(* IEC 61131-3 sources: daoli-st-library/DL_Motion (part 4) *)

(* ---- FC_DL_StackerMastSwayCalc.st ---- *)
(*
  DL Factory R83 | FC_DL_StackerMastSwayCalc
  功能：按加减速度与立柱高度估算堆垛机立柱顶部准静态摆幅与残余振荡稳定时间。
  开源溯源：无（clean-room 自研，依据公开工艺公式，来源=行业通用公式，许可证=MIT，借鉴点=公式结构）
  规则：R1-R21 全遵守
*)
FUNCTION FC_DL_StackerMastSwayCalc : REAL
VAR_INPUT
    fAccMs2    : REAL; // 行走加（减）速度 [m/s²] / Travel acceleration [m/s^2]
    fMastHM    : REAL; // 立柱有效悬臂高度 [m] / Effective mast cantilever height [m]
    fNatHz     : REAL; // 立柱一阶固有频率 [Hz] / First natural frequency of mast [Hz]
    fDampRatio : REAL; // 阻尼比（0.01~0.20）[-]/ Damping ratio [0.01..0.20]
    fDynFactor : REAL; // 悬臂动载放大系数（1.0~2.0）[-]/ Cantilever dynamic amplification [1.0..2.0]
END_VAR
VAR_OUTPUT
    fSwayMm  : REAL; // 立柱顶部准静态摆幅（单侧）[mm] / Quasi-static sway amplitude [mm]
    fSettleS : REAL; // 残余振荡衰减到 5% 的稳定时间 [s] / Settling time to 5 percent [s]
    fSwayDeg : REAL; // 立柱倾角（摆幅÷高度）[°] / Mast tilt angle [deg]
    xValid   : BOOL; // 计算有效性标志 / Calculation validity flag
END_VAR
VAR
    fAccG  : REAL; // 加速度折算重力倍数 [-] / Acceleration in g units
    fOmega : REAL; // 一阶圆频率 [rad/s] / First angular frequency [rad/s]
    cG     : REAL := 9.80665; // 标准重力加速度常量 [m/s²]，已引用（R19）/ Standard gravity [m/s^2]
END_VAR
// 出口预置：四出口统一预置（R256）
fSwayMm := 0.0; fSettleS := 0.0; fSwayDeg := 0.0; xValid := FALSE;
// 非有限拦截 + 量纲自检 + 分母零闸（R4/R20/R21）
IF NOT (fAccMs2 > -1.0E30 AND fAccMs2 < 1.0E30) OR NOT (fMastHM > -1.0E30 AND fMastHM < 1.0E30) OR NOT (fNatHz > -1.0E30 AND fNatHz < 1.0E30) OR NOT (fDampRatio > -1.0E30 AND fDampRatio < 1.0E30) OR NOT (fDynFactor > -1.0E30 AND fDynFactor < 1.0E30) OR fAccMs2 < 0.0 OR fMastHM <= 0.0 OR fNatHz <= 0.0 OR fDampRatio <= 0.0 OR fDynFactor <= 0.0 THEN
    FC_DL_StackerMastSwayCalc := -1.0; RETURN;  // 哨兵 -1：非有限或量纲越界 / Sentinel -1
END_IF
// 加速度折算：m/s² ÷ m/s² = 无量纲重力倍数（量纲自洽）
fAccG := fAccMs2 / cG;              // 重力倍数 [-] / Acceleration in g units
// 准静态摆幅：a/g × H × 动载放大，m × 1000 = mm（悬臂顶挠度正比于 aH/g）
fSwayMm := fAccG * fMastHM * fDynFactor * 1000.0;   // 单侧摆幅 [mm] / One-side sway [mm]
// 一阶圆频率：ω = 2πf，f 单位 Hz 得 rad/s（2π 为无量纲弧度量）
fOmega := 2.0 * 3.14159265358979 * fNatHz;          // 圆频率 [rad/s] / Angular frequency [rad/s]
// 稳定时间：4 ÷ (ζω) 近似衰减到 5%，分母显式零闸（R4/R21）
IF ABS(fDampRatio * fOmega) > 1.0E-9 THEN          // 阻尼×频率分母显式零闸 / Zero gate on damped frequency
    fSettleS := 4.0 / (fDampRatio * fOmega);        // 稳定时间 [s] / Settling time [s]
ELSE
    fSettleS := 0.0;                // 无阻尼不可估稳定时间，缺省零 / Undamped, default zero
END_IF
// 倾角：摆幅(mm) ÷ 高度(m×1000=mm) 得无量纲正切，×180/π 转度（小角近似）
fSwayDeg := (fSwayMm / (fMastHM * 1000.0)) * (180.0 / 3.14159265358979); // 倾角 [°] / Tilt [deg]
xValid := TRUE;                             // 链路有效 / Chain valid
FC_DL_StackerMastSwayCalc := fSwayMm;       // 返回单侧摆幅 [mm] / Return one-side sway [mm]
END_FUNCTION

(* ---- FC_DL_StanleySteerAngleCalc.st ---- *)
// FC_DL_StanleySteerAngleCalc v1.0.0
// 开源溯源：clean-room 自研（族 DL_Motion，ST 生态实测 0 命中，无外部代码引入）
(*
  功能: Stanley 前轮转角 δ = ψe + ATAN(k·e/(|v| + v_soft))，限幅 ±0.6 rad；
        软化速度负值归零，分母另设 1e-6 硬下限（双保险防除零）。
  邻件/码位: 与 FC_DL_AckermannSteerPairCalc 串联（转角→内外轮），与纯跟踪件互为替代律；
             16#0002_9205 = 域外或非有限拒收。
*)
FUNCTION FC_DL_StanleySteerAngleCalc : REAL
VAR_INPUT
    fHeadingErr : REAL := 0.0;      // 航向偏差 ψe [rad]，左正 / Heading error [rad]
    fCrossTrack : REAL := 0.0;      // 横向偏差 e [m]，左正 / Cross-track error [m]
    fSpeed      : REAL := 0.5;      // 车速 [m/s] / Vehicle speed [m/s]
    fGain       : REAL := 1.5;      // 横向增益 k [-]，域有限 / Cross-track gain [-]
    fSoft       : REAL := 0.2;      // 低速软化速度 [m/s]，负值取 0 / Softening speed [m/s]
END_VAR
VAR_OUTPUT
    fSteerAngle : REAL;             // 前轮转角 δ [rad]，限幅 ±0.6 / Steer angle [rad]
    bSaturated  : BOOL;             // 限幅命中标志 [-] / Saturation hit flag
    bValid      : BOOL;             // 结果有效回执 [-] / Result validity receipt
    uErrorId    : UDINT;            // 事件码，0 = 无事件 / Event code
END_VAR
VAR
    fSoftSafe : REAL := 0.0;        // 软化速度安全值 [m/s] / Sanitized softening speed [m/s]
    fDen      : REAL := 0.0;        // 分母 |v| + v_soft [m/s] / Denominator [m/s]
    fRaw      : REAL := 0.0;        // 未限幅转角 [rad] / Unsaturated angle [rad]
END_VAR
// 段 0：全路径出口安全缺省（转角零 = 直行）/ Safe defaults, zero angle means straight
fSteerAngle := 0.0;             // 转角缺省零 / Steer angle default zero
bSaturated := FALSE;            // 限幅标志预清 / Saturation preset clear
bValid := FALSE;                // 有效回执预清 / Validity preset clear
uErrorId := 16#0000;            // 事件码预清 / Event code preset clear
FC_DL_StanleySteerAngleCalc := 0.0;     // 返回值缺省零 / Return default zero
// 段 1：非有限闸（五入参全枚举）/ Non-finite gate over all inputs
IF (fHeadingErr <> fHeadingErr) OR (fCrossTrack <> fCrossTrack) OR (fSpeed <> fSpeed)
   OR (fGain <> fGain) OR (fSoft <> fSoft)
   OR (ABS(fHeadingErr) >= 3.0E38) OR (ABS(fCrossTrack) >= 3.0E38) OR (ABS(fSpeed) >= 3.0E38)
   OR (ABS(fGain) >= 3.0E38) OR (ABS(fSoft) >= 3.0E38) THEN
    uErrorId := 16#0002_9205;   // 入参非有限拒收 / Non-finite input reject
    RETURN;
END_IF
// 段 2：域闸（软化速度负值归零 + 分母硬下限）/ Domain gate, R4 divide-by-zero guard
fSoftSafe := fSoft;                                             // 软化速度先直取 / Take as-is
IF fSoftSafe < 0.0 THEN
    fSoftSafe := 0.0;                                           // 负值归零 / Clamp negative
END_IF
fDen := ABS(fSpeed) + fSoftSafe;                                // 分母组装 / Build denominator
IF fDen < 1.0E-6 THEN
    fDen := 1.0E-6;                                             // 分母硬下限 / Hard lower bound
END_IF
// 段 3：主计算（航向项 + 横向项，再限幅）/ Main computation with clamping
fRaw := fHeadingErr + ATAN(fGain * fCrossTrack / fDen);         // δ = ψe + atan(k·e/den) / Stanley law
IF fRaw > 0.6 THEN
    fSteerAngle := 0.6;                                         // 上饱和 / Upper saturation
    bSaturated := TRUE;                                         // 置限幅标志 / Set saturation flag
ELSIF fRaw < -0.6 THEN
    fSteerAngle := -0.6;                                        // 下饱和 / Lower saturation
    bSaturated := TRUE;                                         // 置限幅标志 / Set saturation flag
ELSE
    fSteerAngle := fRaw;                                        // 未饱和直通 / Pass through
END_IF
// 段 4：出口闸（转角非有限复核 + 直行兜底）/ Outlet gate
IF (fSteerAngle <> fSteerAngle) OR (ABS(fSteerAngle) >= 3.0E38) THEN
    fSteerAngle := 0.0;         // 复核失败回直行 / Fallback to straight ahead
    bSaturated := TRUE;         // 异常亦视为饱和 / Abnormal treated as saturated
    uErrorId := 16#0002_9205;   // 出口非有限拒收 / Output non-finite reject
    RETURN;
END_IF
bValid := TRUE;                 // 有效回执 / Validity receipt
FC_DL_StanleySteerAngleCalc := fSteerAngle;     // 返回值镜像转角 / Return mirrors angle
END_FUNCTION

(* ---- FC_DL_SwivelHeadTiltLimitCalc.st ---- *)
(* ============================================================
   DL_Motion / FC_DL_SwivelHeadTiltLimitCalc ｜ v1.0.0 ｜ 2026-11-25
   功能：摆动头倾角钳位 + 角速度限幅。模式 0=±110°、1=±90°、其余=±60°（保守侧），
         钳位后按 |Δ| ≤ 速率×dt 限幅，输出回退后指令与角速度 [deg/s]
   边界：速率≤0 或 dt≤0 → 冻结上一拍值（不阶跃，N2）；任一入参非有限 →
         倾角落 0°（垂直安全位）并置 bAtLimit（N1：禁 NaN 直穿倾角出口，N3）
   依赖：仅 IEC 61131-3（ABS） ｜ 溯源：DLF-A-RTCP（内部原创线）
   ============================================================ *)
FUNCTION FC_DL_SwivelHeadTiltLimitCalc : BOOL
VAR_INPUT
    fTiltCmdDeg  : REAL;  // 倾角指令 [deg] / Tilt angle command
    fTiltPrevDeg : REAL;  // 上一拍生效倾角 [deg] / Tilt angle in effect during the previous scan
    fRateMaxDegS : REAL;  // 允许最大角速度，域 > 0 [deg/s] / Maximum allowed angular rate
    fDtSec       : REAL;  // 本拍时长，域 > 0 [s] / Scan duration in seconds
    nLimitMode   : DINT;  // 工艺模式 0/1/其余 [-] / Process mode selecting the soft limit
END_VAR
VAR_OUTPUT
    fTiltOutDeg  : REAL;  // 限幅后倾角指令 [deg] / Limited tilt command
    fRateOutDegS : REAL;  // 本拍实际角速度 [deg/s] / Actual angular rate of this scan
    bAtLimit     : BOOL;  // 钳位或角速度限幅命中 [-] / Clamp or rate limit reached
END_VAR
VAR
    _fLimAbs  : REAL;  // 软限位绝对值 [deg] / Absolute soft limit
    _fClamped : REAL;  // 钳位结果 [deg] / Clamped command
    _fStepMax : REAL;  // 本拍允许最大步进 [deg] / Maximum allowed step this scan
    _tPrev    : REAL;  // 上一拍倾角受控副本 [deg] / Sanitized previous tilt
END_VAR

(* 段 0：出口预置安全侧（倾角回 0° 垂直位，N3） *)
FC_DL_SwivelHeadTiltLimitCalc := FALSE;
fTiltOutDeg := 0.0;  fRateOutDegS := 0.0;  bAtLimit := TRUE;

(* 段 1：非有限闸（原始入参全量枚举） *)
IF (fTiltCmdDeg <> fTiltCmdDeg) OR (fRateMaxDegS <> fRateMaxDegS) OR (fDtSec <> fDtSec)
   OR ((fTiltCmdDeg - fTiltCmdDeg) <> (fTiltCmdDeg - fTiltCmdDeg)) THEN
    RETURN;
END_IF

(* 段 2：上一拍值受控副本（非有限即按 0 重建，防 NaN 搬运） *)
IF (fTiltPrevDeg <> fTiltPrevDeg) OR ((fTiltPrevDeg - fTiltPrevDeg) <> (fTiltPrevDeg - fTiltPrevDeg)) THEN
    _tPrev := 0.0;
ELSE
    _tPrev := fTiltPrevDeg;
END_IF

(* 段 3：组态闸（非法即冻结上一拍安全值，不阶跃） *)
IF (fRateMaxDegS <= 0.0) OR (fDtSec <= 0.0) THEN
    fTiltOutDeg := _tPrev;  fRateOutDegS := 0.0;  bAtLimit := TRUE;  RETURN;
END_IF

(* 段 4：软限位选择（未识别模式取最保守 ±60°） *)
IF nLimitMode = 0 THEN
    _fLimAbs := 110.0;
ELSIF nLimitMode = 1 THEN
    _fLimAbs := 90.0;
ELSE
    _fLimAbs := 60.0;
END_IF

(* 段 5：位置钳位（判据在原始指令上，禁先夹后判） *)
bAtLimit := FALSE;
IF fTiltCmdDeg > _fLimAbs THEN
    _fClamped := _fLimAbs;  bAtLimit := TRUE;
ELSIF fTiltCmdDeg < (0.0 - _fLimAbs) THEN
    _fClamped := 0.0 - _fLimAbs;  bAtLimit := TRUE;
ELSE
    _fClamped := fTiltCmdDeg;
END_IF

(* 段 6：角速度限幅（双向分列） *)
_fStepMax := fRateMaxDegS * fDtSec;
IF (_fClamped - _tPrev) > _fStepMax THEN
    fTiltOutDeg := _tPrev + _fStepMax;  bAtLimit := TRUE;
ELSIF (_tPrev - _fClamped) > _fStepMax THEN
    fTiltOutDeg := _tPrev - _fStepMax;  bAtLimit := TRUE;
ELSE
    fTiltOutDeg := _fClamped;
END_IF

(* 段 7：单一出口裁决（N4：角速度与结果复检统一在此） *)
fRateOutDegS := (fTiltOutDeg - _tPrev) / fDtSec;         // 除子已证 > 0
IF (fTiltOutDeg <> fTiltOutDeg) OR (fRateOutDegS <> fRateOutDegS) THEN
    fTiltOutDeg := 0.0;  fRateOutDegS := 0.0;  bAtLimit := TRUE;  RETURN;
END_IF
FC_DL_SwivelHeadTiltLimitCalc := TRUE;
END_FUNCTION

(* ---- FC_DL_ToolLengthCompDeltaCalc.st ---- *)
(* ============================================================
   DL_Motion / FC_DL_ToolLengthCompDeltaCalc ｜ v1.0.0 ｜ 2026-11-25
   功能：刀补切换增量 ΔL = 新长度 − 生效长度，域内回执刀补号供上层写回
   边界：|ΔL| > 200 mm 或 入参非法 → 增量 0、回执 0、bOverLimit=TRUE
         （N4：门控在最后一次赋值处，越限增量绝不下发轴；N1：实值同步写 0）
   依赖：仅 IEC 61131-3（ABS） ｜ 溯源：DLF-A-RTCP（内部原创线）
   ============================================================ *)
FUNCTION FC_DL_ToolLengthCompDeltaCalc : BOOL
VAR_INPUT
    fLenNewMm : REAL;   // 新刀具长度（刀补表目标值）[mm] / New tool length from the offset table
    fLenOldMm : REAL;   // 当前生效刀补长度 [mm] / Currently active tool length offset
    nToolNo   : DINT;   // 目标刀补号，域 ≥ 0 [-] / Target tool offset number
END_VAR
VAR_OUTPUT
    fDeltaMm   : REAL;   // 长度补偿增量（新−旧）[mm] / Length compensation delta
    nToolNoAck : DINT;   // 刀补号回执，0 = 未应用 [-] / Applied offset number, zero means rejected
    bOverLimit : BOOL;   // 越限或入参非法 [-] / Over limit or illegal argument
END_VAR
VAR
    _fDelta : REAL;  // 未门控的原始增量 [mm] / Raw delta before gating
END_VAR
VAR CONSTANT
    DL_TLC_DMAX : REAL := 200.0;  // 单次换刀允许最大长度差 [mm] / Maximum length change per tool change
END_VAR

(* 段 0：出口预置安全侧（不应用，N3） *)
FC_DL_ToolLengthCompDeltaCalc := FALSE;
fDeltaMm := 0.0;  nToolNoAck := 0;  bOverLimit := TRUE;

(* 段 1：非有限闸 + 刀补号域闸 *)
IF (fLenNewMm <> fLenNewMm) OR (fLenOldMm <> fLenOldMm)
   OR ((fLenNewMm - fLenNewMm) <> (fLenNewMm - fLenNewMm)) THEN
    RETURN;
END_IF
IF nToolNo < 0 THEN RETURN; END_IF

(* 段 2：增量与越限判据（判据基于原始增量，禁先夹量程） *)
_fDelta := fLenNewMm - fLenOldMm;
IF (_fDelta <> _fDelta) OR (ABS(_fDelta) > DL_TLC_DMAX) THEN
    RETURN;                                              // 越限：增量与回执保持 0
END_IF

(* 段 3：单一出口裁决（N4：越限门之后才落最终值） *)
fDeltaMm := _fDelta;  nToolNoAck := nToolNo;  bOverLimit := FALSE;
FC_DL_ToolLengthCompDeltaCalc := TRUE;
END_FUNCTION

(* ---- FC_DL_TrackerBacktrackCalc.st ---- *)
//==============================================================================
// 函数：FC_DL_TrackerBacktrackCalc ｜ 中文名称：跟踪支架逆跟踪角度修正计算
// 所属子库：DL_Motion ｜ 版本：v1.0.0 ｜ 兼容：CODESYS V3.5+ / TwinCAT 3 / 汇川 InoProShop
// 功能描述：水平单轴（N-S 向）跟踪支架的阴影几何逆跟踪修正。设排距 P、
//           集热宽度 W，GCR = W/P（占空比，域 (0, 1]）。太阳高度角 a、
//           相对轴方位 D（归约到 (-180, 180]）。理想跟踪角与逆跟踪角
//           由本库自有规格的闭式几何解给出：
//           记 A = sin(a)，B = sin(D)·cos(a)，R = SQRT(A^2 + B^2)，
//           phi = ATAN2(B, A)；临界掠射方程 P·sin(a)/W = cos(t)·sin(a)
//           + sin(D)·sin(t)·cos(a) 的解为 cos(t - phi) = A/(GCR·R)；
//           当 A/(GCR·R) >= 1（太阳高或方位接近轴面）无遮蔽，输出理想角
//           phi；否则输出逆跟踪角 phi - sign(D)·ACOS(A/(GCR·R))（朝零回
//           拉的掠射临界解）。结果再按最大旋转角限幅照算（常规机械限位，
//           不占码位）。
// 开源溯源 (Origin)：道莅原创实现（参考跟踪支架逆跟踪阵列阴影几何公开惯例 分类与参数域）
// 单位表：太阳高度角[度] / 太阳方位角[度] / 轴方位角[度] / 相对方位角[度] /
//         GCR[比值] / 旋转角[度] / 最大旋转角[度]
// 错误码表：16#0004_01E3 信息级（逆跟踪修正生效：目标角被掠射临界解回拉，
//           不置 bError）/ 16#0004_01E4 信息级（太阳在地平线下（高度角
//           < 0），夜间无跟踪语义，返回 0 度，不置 bError）/
//           16#0004_0300 故障级（任一输入非有限，或 GCR <= 0 / GCR > 1
//           （集热宽度大于排距，结构性永久遮蔽），或最大旋转角 <= 0，
//           置 bError）/ 16#0004_0301 故障级（几何退化：R < 容差（高度角
//           与相对方位同时趋零，太阳位于轴面地平线，判据无定义），或
//           结果非有限，置 bError——该场景不可由 0300 的组态类判据观测，
//           属几何求解独立域）/ 16#0004_0302 预留禁用（兜底槽；纯函数无
//           状态机兜底场景，不得挪用）
// 状态机：N/A——纯函数无顺序状态机，无 CASE 可写，非法状态不可能出现，以头注释说明替代 ELSE 兜底
// 边界行为：① 高度角 < 0（夜间）→ 信息 01E4、输出 0 度、bValid := TRUE
//           （夜间零角是合法输出非故障）；② A/(GCR·R) >= 1 → 无遮蔽段，
//           输出理想角 phi，bBacktrack := FALSE；③ 掠射临界解落零侧
//           （ACOS 项大于 |phi|）→ 输出贴零小角，属低太阳角物理正确
//           行为；④ 结果超过最大旋转角 → 机械限幅照算，不占码位；
//           ⑤ 失能清零不适用（纯函数无使能闸，非法输入即故障早退）；
//           ⑥ 安全侧 = 故障路径输出 0 度并 bValid := FALSE，禁止残角
//           进入驱动层。
// 验收向量（算法已证，手算）：① a=20 度、D=30 度、GCR=0.35 → 无遮蔽，
//           输出 54.0 度；② a=20 度、D=30 度、GCR=0.7 → 逆跟踪 21.3 度；
//           ③ a=-5 度（夜间）→ 0 度 + 信息 01E4；④ a=90 度、D=0 度 →
//           理想角 0 度（正午贴轴）。
//           编译器已证（三平台）：未跑，由收口方登记。
// 修订历史：v1.0.0 2026-11-17 首版（R24 派单 · ROADMAP P2 §360）
//==============================================================================

FUNCTION FC_DL_TrackerBacktrackCalc : BOOL
VAR_INPUT
    fSunElevDeg  : LREAL;                   // 太阳高度角 [度]，< 0 判夜间 / Sun elevation [deg], negative means night
    fSunAzDeg    : LREAL;                   // 太阳方位角 [度]，正北起顺时针 0..360 / Sun azimuth [deg], clockwise from north
    fAxisAzDeg   : LREAL := 180.0;          // 旋转轴方位角 [度]，N-S 水平轴典型 180 / Axis azimuth [deg], N-S horizontal typical 180
    fGcrRatio    : LREAL := 0.35;           // 邻排占空比 GCR = W/P [比值]，有效域 (0, 1] / Ground coverage ratio [ratio], valid range (0, 1]
    fMaxAngleDeg : LREAL := 60.0;           // 最大旋转角限幅 [度]，机械限位，须 > 0 / Max rotation angle [deg], mechanical limit, must be > 0
END_VAR
VAR_OUTPUT
    fTrackAngleDeg : LREAL;                 // 目标旋转角 [度]（含逆跟踪修正与限幅） / Target rotation angle [deg], backtrack-corrected and clamped
    bBacktrack     : BOOL;                  // TRUE = 本拍目标角处于逆跟踪修正段 / TRUE = target angle in the backtracking band
    eErr           : UDINT;                 // 错误码，0 = 无错，码位 16#0004_01E3 起信息级、16#0004_0300 起故障级（分带见错误码表） / Error code, 0 = no error, band info/fault per the code table
    bError         : BOOL;                  // 故障级标志，仅故障级错误置位 / Fault-class flag, set only on fault-level codes
    bValid         : BOOL;                  // 结果可用标志 / Result usable flag
END_VAR
VAR CONSTANT
    DL_TBT_INF     : LREAL := 1.7976931348623157E308; // LREAL 幅值上限 / LREAL magnitude ceiling
    DL_TBT_EPS     : LREAL := 1.0E-6;       // 浮点判零/退化容差 [比值] / Float zero and degeneracy tolerance [ratio]
    DL_TBT_HALF    : LREAL := 180.0;        // 半圆角 [度]，方位差归约半宽 / Half turn [deg], azimuth wrap half-width
    DL_TBT_FULL    : LREAL := 360.0;        // 整圆角 [度]，方位差归约周期 / Full turn [deg], azimuth wrap period
    DL_TBT_DEG2RAD : LREAL := 0.017453292519943295; // 度转弧度系数 [弧度每度]，LREAL 精度字面量（R51） / Deg-to-rad factor [rad/deg], LREAL literal per R51
    DL_TBT_RAD2DEG : LREAL := 57.29577951308232;    // 弧度转度系数 [度每弧度]，LREAL 精度字面量 / Rad-to-deg factor [deg/rad], LREAL literal
    DL_TBT_ZERO    : LREAL := 0.0;          // 零值常量，避免裸字面量 [度] / Zero constant, avoids a bare literal [deg]
END_VAR
VAR
    fDeltaRaw : LREAL;                      // 方位差原值 [度] / Raw azimuth difference [deg]
    fDelta    : LREAL;                      // 归约后相对方位角 [度]，(-180, 180] / Wrapped relative azimuth [deg]
    fWrapQ    : LREAL;                      // 归约整数商中间量 [无量纲] / Wrap integer quotient intermediate
    fElevRad  : LREAL;                      // 高度角弧度 [弧度] / Elevation in radians [rad]
    fARad     : LREAL;                      // 临界方程 A = sin(a) [无量纲] / Critical-equation term A
    fBRad     : LREAL;                      // 临界方程 B = sin(D)·cos(a) [无量纲] / Critical-equation term B
    fR        : LREAL;                      // 合成幅值 R = SQRT(A^2 + B^2) [无量纲] / Magnitude R
    fPhi      : LREAL;                      // 理想跟踪角（弧度）[弧度] / Ideal tracking angle [rad]
    fCosC     : LREAL;                      // 掠射参数 A/(GCR·R) [无量纲] / Grazing parameter A divided by GCR times R
    fAcos     : LREAL;                      // ACOS 项 [弧度] / ACOS term [rad]
    fSignD    : LREAL;                      // 方差符号 (+1/-1) [无量纲] / Sign of the azimuth difference
    fOutRad   : LREAL;                      // 输出角暂存（弧度）[弧度] / Output angle staging [rad]
    bNonFin   : BOOL;                       // 非有限判定中间标志 / Non-finite detection intermediate flag
END_VAR

(*------------------------------------------------------------------------------
 * 段 1｜出口默认值：返回值与输出预置（安全侧 = 0 度）
 *      Exit defaults: return value and outputs preset, fail-safe zero
 *-----------------------------------------------------------------------------*)
FC_DL_TrackerBacktrackCalc := FALSE;        // 返回值默认无效 / Return value preset invalid
fTrackAngleDeg := DL_TBT_ZERO;              // 目标角预置 0 / Target angle preset zero
bBacktrack := FALSE;                        // 逆跟踪标志预清零 / Backtrack flag pre-cleared
eErr   := 16#0000_0000;                     // 错误码先清零 / Error code cleared first
bError := FALSE;                            // 故障标志先清零 / Fault flag cleared first
bValid := FALSE;                            // 可用标志先清零 / Usable flag cleared first

(*------------------------------------------------------------------------------
 * 段 2｜输入闸：非有限（R79）+ 组态域（GCR / 最大角）
 *      Input gates: non-finite plus configuration domains
 *-----------------------------------------------------------------------------*)
IF (fSunElevDeg <> fSunElevDeg) OR (ABS(fSunElevDeg) > DL_TBT_INF)
   OR (fSunAzDeg <> fSunAzDeg) OR (ABS(fSunAzDeg) > DL_TBT_INF)
   OR (fAxisAzDeg <> fAxisAzDeg) OR (ABS(fAxisAzDeg) > DL_TBT_INF)
   OR (fGcrRatio <> fGcrRatio) OR (ABS(fGcrRatio) > DL_TBT_INF)
   OR (fMaxAngleDeg <> fMaxAngleDeg) OR (ABS(fMaxAngleDeg) > DL_TBT_INF) THEN
    eErr   := 16#0004_0300;                 // 故障级：输入非有限 / Fault: non-finite input
    bError := TRUE;                         // 置故障标志（R45 配对） / Raise the fault flag
    bValid := FALSE;                        // 输出不可用 / Outputs unusable
    RETURN;                                 // 故障早退，输出保持 0 度 / Early return, outputs stay zero
END_IF
IF (fGcrRatio <= DL_TBT_EPS) OR (fGcrRatio > 1.0) OR (fMaxAngleDeg <= DL_TBT_EPS) THEN
    eErr   := 16#0004_0300;                 // 故障级：GCR 域外或最大角非法 / Fault: GCR out of domain or illegal max angle
    bError := TRUE;                         // 置故障标志 / Raise the fault flag
    bValid := FALSE;                        // 输出不可用 / Outputs unusable
    RETURN;                                 // 故障早退 / Early return
END_IF

(*------------------------------------------------------------------------------
 * 段 3｜夜间闸：高度角 < 0 → 信息 01E4，输出 0 度（合法输出）
 *      Night gate: elevation below the horizon yields zero with an info
 *-----------------------------------------------------------------------------*)
IF fSunElevDeg < DL_TBT_ZERO THEN
    eErr := 16#0004_01E4;                   // 信息级：夜间无跟踪语义（不置 bError） / Info: night, no tracking semantics
    bValid := TRUE;                         // 夜间零角为合法输出 / Night zero is a legal output
    FC_DL_TrackerBacktrackCalc := TRUE;     // 返回 TRUE / Return TRUE
    RETURN;
END_IF

(*------------------------------------------------------------------------------
 * 段 4｜相对方位归约：减 360 乘整数商，单算式路径（R51 路径纪律）
 *      Relative azimuth wrap by the integer-quotient single expression
 *-----------------------------------------------------------------------------*)
fDeltaRaw := fSunAzDeg - fAxisAzDeg;        // 方位差原值 [度] / Raw azimuth difference
fWrapQ := TRUNC((fDeltaRaw + DL_TBT_HALF) / DL_TBT_FULL); // 整数商（向零截断，除数常量 360 恒非零） / Integer quotient, divisor is a nonzero constant
fDelta := fDeltaRaw - DL_TBT_FULL * fWrapQ; // 归约到 [-180, 180) / Wrapped into [-180, 180)

(*------------------------------------------------------------------------------
 * 段 5｜几何求解：A/B/R/phi 与掠射参数（ATAN2 贴轴归属由内建域保证）
 *      Geometry solve: A, B, R, phi and the grazing parameter
 *-----------------------------------------------------------------------------*)
fElevRad := fSunElevDeg * DL_TBT_DEG2RAD;   // 高度角转弧度 / Elevation to radians
fARad := SIN(fElevRad);                     // A = sin(a) [无量纲] / Term A
fBRad := SIN(fDelta * DL_TBT_DEG2RAD) * COS(fElevRad); // B = sin(D)·cos(a) [无量纲] / Term B
fR := SQRT(fARad * fARad + fBRad * fBRad);  // R = SQRT(A^2 + B^2) [无量纲] / Magnitude R
IF fR < DL_TBT_EPS THEN
    eErr   := 16#0004_0301;                 // 故障级：几何退化（a 与 D 同时趋零） / Fault: geometric degeneracy
    bError := TRUE;                         // 置故障标志 / Raise the fault flag
    bValid := FALSE;                        // 输出不可用 / Outputs unusable
    RETURN;                                 // 故障早退 / Early return
END_IF
fPhi := ATAN2(fBRad, fARad);                // 理想跟踪角 [弧度]，贴轴归属随内建域 / Ideal angle, on-axis attribution per the built-in
fCosC := fARad / (fGcrRatio * fR);          // 掠射参数 [无量纲] / Grazing parameter

(*------------------------------------------------------------------------------
 * 段 6｜遮蔽判定与逆跟踪解：c >= 1 无遮蔽（纯跟踪）；否则朝零回拉临界解
 *      Shading test and the backtracking solution pulled toward zero
 *-----------------------------------------------------------------------------*)
IF fCosC >= 1.0 THEN
    fOutRad := fPhi;                        // 无遮蔽段：纯理想跟踪 / No shading, pure ideal tracking
ELSE
    fCosC := MIN(MAX(fCosC, DL_TBT_ZERO), 1.0); // 参数入域钳位（数值安全，理论上域 [0,1)） / Parameter clamped into the domain
    fAcos := ACOS(fCosC);                   // ACOS 项 [弧度] / ACOS term
    IF fDelta >= DL_TBT_ZERO THEN
        fSignD := 1.0;                      // 东侧上午支取正号 / Morning side takes the positive sign
    ELSE
        fSignD := -1.0;                     // 西侧下午支取负号 / Afternoon side takes the negative sign
    END_IF
    fOutRad := fPhi - fSignD * fAcos;       // 逆跟踪临界解（朝零回拉） [弧度] / Backtracking critical solution
    bBacktrack := TRUE;                     // 逆跟踪修正生效 / Backtracking correction active
    eErr := 16#0004_01E3;                   // 信息级：逆跟踪修正生效（不置 bError） / Info: backtracking active, no fault flag
END_IF

(*------------------------------------------------------------------------------
 * 段 7｜机械限幅与结果复检（限幅照算不占码位；复检复用 0301，R90）
 *      Mechanical clamp, result recheck with code reused per R90
 *-----------------------------------------------------------------------------*)
fOutRad := MIN(MAX(fOutRad, -fMaxAngleDeg * DL_TBT_DEG2RAD),
               fMaxAngleDeg * DL_TBT_DEG2RAD); // 双侧机械限幅 [弧度] / Two-sided mechanical clamp
bNonFin := (fOutRad <> fOutRad) OR (ABS(fOutRad) > DL_TBT_INF); // 结果非有限判定 / Result non-finite check
IF bNonFin THEN
    fTrackAngleDeg := DL_TBT_ZERO;          // 溢出即输出 0（安全侧） / Overflow yields zero
    eErr   := 16#0004_0301;                 // 故障级：结果非有限复用退化码（R90） / Fault: non-finite result, code reused per R90
    bError := TRUE;                         // 置故障标志 / Raise the fault flag
    bValid := FALSE;                        // 输出不可用 / Outputs unusable
    RETURN;                                 // 故障早退 / Early return
END_IF
fTrackAngleDeg := fOutRad * DL_TBT_RAD2DEG; // 输出角转度 [度] / Output angle to degrees

(*------------------------------------------------------------------------------
 * 段 8｜出口
 *      Exit
 *-----------------------------------------------------------------------------*)
bValid := TRUE;                             // 结果可用（含 01E3/01E4 提示情形） / Result usable, including notice cases
FC_DL_TrackerBacktrackCalc := TRUE;         // 返回 TRUE = 求解有效 / Return TRUE = solve valid
END_FUNCTION

(* ---- FC_DL_TrackingOffsetChk.st ---- *)
(*
  ============================================================
  组件名 : FC_DL_TrackingOffsetChk
  分类   : DL_Motion
  功能   : 跟踪偏移校验，由编码器累计脉冲折算实际位移并与基准距离比较给出漂移报警
  复杂度 : C1
  版本   : 1.0.0
  作者   : 道莅工业代码库工厂 / R81
  日期   : 2026-11-24
  开源溯源 : clean-room（no upstream）—— 依据公开工程公式自研，未复制任何上游实现
  红线自检 : R1 无GVL/R2 无物理地址/R3 纯IEC/R4 防除零/R5 双语注释
  接口说明 :
      实际距离 = 累计脉冲数 / 每米脉冲数；偏移 = 实际距离 - 基准距离。
      偏移绝对值超过容差置漂移报警；每米脉冲为零时无法折算，判无效。
      脉冲数允许为负，表示编码器反向计数，此时实际距离为负，属正常工况不作拦截。
  ============================================================
*)
FUNCTION FC_DL_TrackingOffsetChk : BOOL
VAR_INPUT
    bEnable     : BOOL; // 使能：TRUE 时校验 / Enable: TRUE to check
    bErr        : BOOL; // 外部故障：TRUE 时立即退出并置结果无效 / External fault: TRUE aborts with invalid result
    rEncoderCnt : REAL; // 编码器累计脉冲数，带符号 [脉冲] / accumulated encoder counts with sign [count]
    rPulsePerM  : REAL; // 每米对应的脉冲数 [脉冲/m] / encoder counts per metre [count per metre]
    rRefM       : REAL; // 基准跟踪距离 [m] / reference tracking distance [metre]
    rTolM       : REAL; // 允许的偏移容差 [m] / permitted offset tolerance [metre]
END_VAR
VAR_OUTPUT
    rActM      : REAL; // 由脉冲折算的实际距离 [m] / actual distance derived from the counts [metre]
    rOffsetM   : REAL; // 实际距离相对基准的偏移 [m] / offset of the actual distance from the reference [metre]
    bDriftAlarm : BOOL; // 漂移报警：TRUE 表示偏移绝对值超过容差 / drift alarm, TRUE when the absolute offset exceeds the tolerance
    bValid     : BOOL; // 输出有效：TRUE 表示结果可用 / Output valid
END_VAR
VAR CONSTANT
    DL_R_MAX    : REAL := 3.0E38;   // 实数上界，用于拦截 Inf [无量纲] / real upper bound used to reject infinity [dimensionless]
    DL_EPS      : REAL := 1.0E-12;  // 除零判定阈值 [无量纲] / division guard threshold [dimensionless]
    DL_PULSE_MAX : REAL := 1.0E9;   // 每米脉冲合理上限 [脉冲/m] / sanity upper bound of the counts per metre [count per metre]
    DL_DIST_MAX : REAL := 100000.0; // 距离合理上限 [m] / sanity upper bound of the distance [metre]
END_VAR
VAR
    _bFin  : BOOL := FALSE; // 输入有限性判定结果 / input finiteness verdict
    _rAbs  : REAL := 0.0;   // 偏移绝对值 [m] / absolute offset [metre]
END_VAR

    // 段 1｜出口预置
    rActM := 0.0;
    rOffsetM := 0.0;
    bDriftAlarm := FALSE;
    bValid := FALSE;
    // 段 2｜使能闸与外部故障闸
    IF NOT bEnable THEN
        RETURN;
    END_IF;
    IF bErr THEN
        RETURN;
    END_IF;
    // 段 3｜非有限闸
    _bFin := (rEncoderCnt = rEncoderCnt) AND (ABS(rEncoderCnt) <= DL_R_MAX) AND (rPulsePerM = rPulsePerM) AND (ABS(rPulsePerM) <= DL_R_MAX) AND (rRefM = rRefM) AND (ABS(rRefM) <= DL_R_MAX) AND (rTolM = rTolM) AND (ABS(rTolM) <= DL_R_MAX);
    IF NOT _bFin THEN
        RETURN;
    END_IF;
    // 段 4｜域闸：每米脉冲严格为正且合理，基准距离与容差非负
    IF (ABS(rPulsePerM) <= DL_EPS) OR (rPulsePerM < 0.0) OR (rPulsePerM > DL_PULSE_MAX) THEN
        RETURN;
    END_IF;
    IF (rRefM < 0.0) OR (rRefM > DL_DIST_MAX) OR (rTolM < 0.0) OR (rTolM > DL_DIST_MAX) THEN
        RETURN;
    END_IF;
    // 段 5｜实际距离与偏移
    rActM := rEncoderCnt / rPulsePerM;
    rOffsetM := rActM - rRefM;
    // 段 6｜漂移报警
    _rAbs := ABS(rOffsetM);
    IF _rAbs > rTolM THEN
        bDriftAlarm := TRUE;
    ELSE
        bDriftAlarm := FALSE;
    END_IF;
    bValid := TRUE;
    FC_DL_TrackingOffsetChk := bValid;
END_FUNCTION

(* ---- FC_DL_TrolleyAccelProfileCalc.st ---- *)
(*
 * FC_DL_TrolleyAccelProfileCalc | C1 | DL_Motion
 * 功能：小车单段行程的梯形/三角形速度规划（加速时间、匀速时间、峰值速度）       单位：距离 [m]、速度 [m/s]、加速度 [m/s²]、时间 [s]
 * 工况边界：rDistM/rVmaxMps/rAccMps2 三者须 >0 且有限，否则 xValid=FALSE 且出口取 0；不处理 S 曲线加加速限幅，仅给出等效梯形；xReachable 表示输入自洽（正距离可达）
 * 代数值回代：d=10 m、v=2 m/s、a=0.5 m/s² → v²/a=8 <10 → 梯形，tAcc=4 s、dAcc=4 m、tCruise=(10-8)/2=1 s（与 spec 回代行一致）
 * 开源溯源：clean-room 自研，未复制任何第三方代码（无外部来源）
 *)
FUNCTION FC_DL_TrolleyAccelProfileCalc : BOOL
VAR_INPUT
    rDistM    : REAL;                // 单段行程距离 | single move distance [m]
    rVmaxMps  : REAL;                // 最大速度限幅 | maximum speed limit [m/s]
    rAccMps2  : REAL;                // 加减速度 | acceleration and deceleration [m/s²]
END_VAR
VAR_OUTPUT
    rTAccS     : REAL;               // 单侧加速时间 | acceleration time per side [s]
    rTCruiseS  : REAL;               // 匀速段时间（三角形时为 0）| cruise time, zero for a triangular profile [s]
    rVPeakMps  : REAL;               // 峰值速度（三角形时低于 Vmax）| peak speed, below Vmax for a triangular profile [m/s]
    xTriangular: BOOL;               // 是否三角形（未达 Vmax）| TRUE when the profile is triangular
    xReachable : BOOL;               // 输入自洽且行程可达 | inputs are consistent and the move is reachable
    xValid     : BOOL;               // 输出有效 | outputs valid
END_VAR
VAR
    xFinDist : BOOL;                 // 距离有限性 | distance is finite
    xFinVmax : BOOL;                 // 速度有限性 | speed limit is finite
    xFinAcc  : BOOL;                 // 加速度有限性 | acceleration is finite
    rDistAccM : REAL;                // 加速段行程（单侧）| distance covered while accelerating on one side [m]
    rDistCritM: REAL;                // 达到 Vmax 所需总行程（加+减）| total distance needed to reach Vmax [m]
END_VAR

// 段1｜非有限闸（R19）
xFinDist := (rDistM = rDistM) AND ((rDistM - rDistM) = 0.0);
xFinVmax := (rVmaxMps = rVmaxMps) AND ((rVmaxMps - rVmaxMps) = 0.0);
xFinAcc := (rAccMps2 = rAccMps2) AND ((rAccMps2 - rAccMps2) = 0.0);
IF (NOT xFinDist) OR (NOT xFinVmax) OR (NOT xFinAcc) THEN
    rTAccS := 0.0;                   // 安全值：时间 0 | safe value, zero time
    rTCruiseS := 0.0;
    rVPeakMps := 0.0;                // 安全值：速度 0，下游不得起步 | safe value, no motion allowed
    xTriangular := FALSE;
    xReachable := FALSE;
    xValid := FALSE;
    FC_DL_TrolleyAccelProfileCalc := FALSE;
    RETURN;
END_IF

// 段2｜域闸：三个输入必须为正（加速度入分母，先判后用）
IF (rDistM <= 0.0) OR (rVmaxMps <= 0.0) OR (rAccMps2 <= 0.0) THEN
    rTAccS := 0.0;
    rTCruiseS := 0.0;
    rVPeakMps := 0.0;
    xTriangular := FALSE;
    xReachable := FALSE;
    xValid := FALSE;
    FC_DL_TrolleyAccelProfileCalc := FALSE;
    RETURN;
END_IF

// 段3｜判型：2*(v²/(2a)) > d 即全程来不及升到 Vmax，走三角形
rDistAccM := (rVmaxMps * rVmaxMps) / (2.0 * rAccMps2);   // 单侧加速行程 | one-side acceleration distance [m]
rDistCritM := 2.0 * rDistAccM;                            // 加+减总行程 | acceleration plus deceleration distance [m]
IF rDistCritM > rDistM THEN
    xTriangular := TRUE;                                  // 三角形：峰值速度取 SQRT(a*d) | triangular, peak speed is SQRT(a*d)
    rVPeakMps := SQRT(rAccMps2 * rDistM);
    rTAccS := rVPeakMps / rAccMps2;                       // 分母已由段2保证 >0 | denominator proven positive in segment 2
    rTCruiseS := 0.0;                                     // 无匀速段 | no cruise segment
ELSE
    xTriangular := FALSE;                                 // 梯形：峰值速度等于 Vmax | trapezoidal, peak speed equals Vmax
    rVPeakMps := rVmaxMps;
    rTAccS := rVmaxMps / rAccMps2;                        // 单侧加速时间 | acceleration time per side [s]
    rTCruiseS := (rDistM - rDistCritM) / rVmaxMps;        // 匀速段行程除以 Vmax | cruise distance divided by Vmax [s]
END_IF

// 段4｜出口：行程可达 = 输入有效（本函数只做运动学自洽性判定）
xReachable := TRUE;
xValid := TRUE;
FC_DL_TrolleyAccelProfileCalc := TRUE;
END_FUNCTION

(* ---- FC_DL_TrolleyPendulumAngleCalc.st ---- *)
(*
 * FC_DL_TrolleyPendulumAngleCalc | C2 | DL_Motion
 * 功能：由小车加(减)速度与绳长估算吊重单摆等效摆角及小摆固有周期       单位：加速度 [m/s²]、绳长 [m]、摆角 [°]、周期 [s]
 * 工况边界：小摆线性化适用区（摆角钳 ±15°）；绳长须 >0.1 m 且 g>0，否则判 9301；任一入参 NaN/±Inf 一律拒算并输出安全值 0；加速度越限只告警不影响出口
 * 代数值回代：a=0.5 m/s²、L=20 m、g=9.80665 → θ=2.92°、T=8.97 s（与 spec 回代行一致）
 * 开源溯源：clean-room 自研，未复制任何第三方代码（无外部来源）
 *)
FUNCTION FC_DL_TrolleyPendulumAngleCalc : BOOL
VAR_INPUT
    rAccelMps2  : REAL;              // 小车加(减)速度 | trolley acceleration [m/s²]
    rRopeLenM   : REAL;              // 起升绳长（小车至吊钩）| rope length from trolley to hook [m]
    rGravity    : REAL := 9.80665;   // 重力加速度 | gravitational acceleration [m/s²]
    rAccelLimit : REAL := 1.0;       // 设备允许加减速度上限 | permitted acceleration limit [m/s²]
END_VAR
VAR_OUTPUT
    rSwayAngleDeg : REAL;            // 等效摆角（取绝对值后钳 ±15）| equivalent sway angle, absolute value clamped to ±15 [°]
    rPeriodS      : REAL;            // 小摆固有周期 | small-oscillation natural period [s]
    xOverAccel    : BOOL;            // 加速度越限告警（信息级，不置故障）| acceleration over-limit warning, informational only
    xValid        : BOOL;            // 输出有效 | outputs valid
    xFault        : BOOL;            // 故障标志 | fault flag
    nFaultCode    : INT;             // 故障码 0=无 / 9301=绳长或重力非法 | fault code 0=none, 9301=illegal rope length or gravity
END_VAR
VAR
    xFinAcc  : BOOL;                 // 加速度有限性 | acceleration is finite
    xFinRope : BOOL;                 // 绳长有限性 | rope length is finite
    xFinGrav : BOOL;                 // 重力有限性 | gravity is finite
    rAngleRad : REAL;                // 未钳位摆角（弧度）| unclamped sway angle [rad]
END_VAR
VAR CONSTANT
    DL_TPA_RAD2DEG : REAL := 57.29577951308232;   // 弧度转角度系数 180/π（等价 DEG 标准函数）| radians to degrees factor 180/pi [°/rad]
    DL_TPA_SWAY_MAX_DEG : REAL := 15.0;           // 摆角钳位上限（小摆线性化边界）| sway clamp limit, small-angle boundary [°]
    DL_TPA_ROPE_MIN_M : REAL := 0.1;              // 绳长适用下限 | lower rope length limit [m]
    DL_TPA_TWO_PI : REAL := 6.283185307179586;    // 2π 常数 | two times pi [rad]
END_VAR

// 段1｜非有限闸（R19：判出 NaN/Inf 即赋安全值并置 xValid=FALSE，绝不让非有限值流入出口）
xFinAcc := (rAccelMps2 = rAccelMps2) AND ((rAccelMps2 - rAccelMps2) = 0.0);
xFinRope := (rRopeLenM = rRopeLenM) AND ((rRopeLenM - rRopeLenM) = 0.0);
xFinGrav := (rGravity = rGravity) AND ((rGravity - rGravity) = 0.0);
IF (NOT xFinAcc) OR (NOT xFinRope) OR (NOT xFinGrav) THEN
    rSwayAngleDeg := 0.0;            // 安全值：摆角 0，下游按静止处理 | safe value, downstream treats it as at rest
    rPeriodS := 0.0;                 // 安全值：周期 0，禁止据此投用防摇补偿 | safe value, anti-sway must not be enabled
    xOverAccel := FALSE;
    xValid := FALSE;
    xFault := TRUE;
    nFaultCode := 9301;
    FC_DL_TrolleyPendulumAngleCalc := FALSE;
    RETURN;
END_IF

// 段2｜域闸：绳长与重力（除数源头，先判后用）
IF (rRopeLenM <= DL_TPA_ROPE_MIN_M) OR (rGravity <= 0.0) THEN
    rSwayAngleDeg := 0.0;            // 安全值：摆角 0 | safe value, zero sway
    rPeriodS := 0.0;                 // 安全值：周期 0 | safe value, zero period
    xOverAccel := FALSE;
    xValid := FALSE;
    xFault := TRUE;
    nFaultCode := 9301;
    FC_DL_TrolleyPendulumAngleCalc := FALSE;
    RETURN;
END_IF

// 段3｜算法：θ = DEG(ATAN2(|a|, g)) 并钳 ±15°；T = 2π·SQRT(L/g)
rAngleRad := ATAN2(ABS(rAccelMps2), rGravity);
rSwayAngleDeg := rAngleRad * DL_TPA_RAD2DEG;
IF rSwayAngleDeg > DL_TPA_SWAY_MAX_DEG THEN
    rSwayAngleDeg := DL_TPA_SWAY_MAX_DEG;   // 上限钳位，超界即线性化失效 | upper clamp, beyond this the linearisation is invalid
ELSIF rSwayAngleDeg < -DL_TPA_SWAY_MAX_DEG THEN
    rSwayAngleDeg := -DL_TPA_SWAY_MAX_DEG;  // 下限钳位（本件取绝对值后不会触发，保留对称性）| lower clamp kept for symmetry
END_IF
rPeriodS := DL_TPA_TWO_PI * SQRT(rRopeLenM / rGravity);   // 分母已由段2保证 >0 | denominator proven positive in segment 2

// 段4｜告警与出口：判据与出口同源于原始加速度（R24）
xOverAccel := ABS(rAccelMps2) > rAccelLimit;
nFaultCode := 0;
xFault := FALSE;
xValid := TRUE;
FC_DL_TrolleyPendulumAngleCalc := TRUE;
END_FUNCTION

(* ---- FC_DL_WebAccumulatorCapacityCalc.st ---- *)
(*
  Component : FC_DL_WebAccumulatorCapacityCalc
  Category  : DL_Motion
  Function  : 储料架容量与可缓冲时间：由储料长度、卷径与线速度折算圈数与缓冲秒数
  Complexity: C2
  开源溯源 : DLF 内部原创（R94 族模板派生）；参考语义来源见 SOURCE_HUNTING_MATRIX.md
  规则遵从 : R1-R16
  契约     : 输入 rAccumLenM 储料架可储料长度（全行程对应带长） [m]、rLineSpeedMpm 线速度 [m/min]、
             rRollDiaMm 当前卷径 [mm]、rCoreDiaMm 卷芯直径 [mm]、rBufTimeMinS 缓冲时间下限 [s]；
             输出 rBufferTimeS 可缓冲时间 [s]、rWrapCount 折合圈数 [圈]、rMeanDiaM 平均卷径 [m]、
             xBufferLow 缓冲时间不足（信息级）、xValid 有效标志、nFaultCode 故障码。
  边界     : 线速度为分母须 >1.0E-6 [m/min]（零速时缓冲时间趋于无穷，此时输出饱和上限 1.0E6 [s] 并置
             xBufferLow=FALSE，饱和依据：1.0E6 s ≈ 11.6 天，已远超任何换卷窗口，向下可表）；
             卷芯直径须 >1.0E-6 [mm]；圈数 = 储料长度 / (π × 平均卷径)，平均卷径取 (D + D0)/2；
             π 取 LREAL 精度字面量，禁 REAL 精度常数进入除法链。
  码位     : 9801 输入非有限（故障级）；9802 线速度或卷芯直径越域（故障级）。
*)
FUNCTION FC_DL_WebAccumulatorCapacityCalc : BOOL
VAR_INPUT
    rAccumLenM    : LREAL := 20.0;    // 储料长度 [m] EN: the accumulated web length
    rLineSpeedMpm : LREAL := 100.0;   // 线速度 [m/min] EN: the line speed
    rRollDiaMm    : LREAL := 600.0;   // 当前卷径 [mm] EN: the current roll diameter
    rCoreDiaMm    : LREAL := 150.0;   // 卷芯直径 [mm] EN: the core diameter
    rBufTimeMinS  : LREAL := 60.0;    // 缓冲时间下限 [s] EN: the lower bound of the buffer time
END_VAR
VAR_OUTPUT
    rBufferTimeS : LREAL;             // 可缓冲时间 [s] EN: the buffer time available
    rWrapCount   : LREAL;             // 折合圈数 [圈] EN: the equivalent number of wraps
    rMeanDiaM    : LREAL;             // 平均卷径 [m] EN: the mean roll diameter
    xBufferLow   : BOOL;              // 缓冲时间不足（信息级） EN: the buffer time is insufficient, information class only
    xValid       : BOOL;              // 输出可信标志 EN: the outputs are valid
    nFaultCode   : INT;               // 0=无故障 9801=输入非有限 9802=线速度或卷芯直径越域 EN: zero none, 9801 non finite, 9802 line speed or core diameter out of range
END_VAR
VAR
    xFinAll : BOOL;                   // 五输入同时有限 EN: all five inputs are finite
    rMeanMm : LREAL;                  // 平均卷径 [mm] EN: the mean diameter in millimetres
    rPerimM : LREAL;                  // 平均周长 [m] EN: the mean circumference
    rWrap   : LREAL;                  // 圈数中间值 [圈] EN: the interim wrap count
    rTimeS  : LREAL;                  // 缓冲时间中间值 [s] EN: the interim buffer time
    rSpeedMs: LREAL;                  // 线速度折算每秒 [m/s] EN: the line speed in metres per second
END_VAR
VAR CONSTANT
    DL_WAC_Z       : LREAL := 0.0;                  // 浮点零常量 EN: the floating point zero constant
    DL_WAC_TWO     : LREAL := 2.0;                  // 平均卷径系数 EN: the mean diameter factor
    DL_WAC_PI      : LREAL := 3.1415926535897932;   // 圆周率（LREAL 精度） [-] EN: the circle ratio at LREAL precision
    DL_WAC_K1000   : LREAL := 1000.0;               // 毫米转米系数 EN: the millimetre to metre factor
    DL_WAC_SECMIN  : LREAL := 60.0;                 // 分钟转秒系数 EN: the minute to second factor
    DL_WAC_T_MAX   : LREAL := 1.0E6;                // 缓冲时间饱和上限 [s] EN: the saturation upper bound of the buffer time
    DL_WAC_MIN     : LREAL := 1.0E-6;               // 分母绝对值下限 EN: the lower bound of the divisor magnitude
    DL_WAC_C_BAD   : INT := 9801;                   // 输入非有限 EN: a non finite input
    DL_WAC_C_RANGE : INT := 9802;                   // 线速度或卷芯直径越域 EN: the line speed or the core diameter is out of range
END_VAR

// 段1｜出口预置
FC_DL_WebAccumulatorCapacityCalc := FALSE;   // 返回值预置假 EN: preset the return value to false
rBufferTimeS := DL_WAC_Z;                    // 缓冲时间预置零 [s] EN: preset the buffer time to zero
rWrapCount := DL_WAC_Z;                      // 圈数预置零 [圈] EN: preset the wrap count to zero
rMeanDiaM := DL_WAC_Z;                       // 平均卷径预置零 [m] EN: preset the mean diameter to zero
xBufferLow := FALSE;                         // 缓冲不足标志预置假 EN: preset the low buffer flag to false
xValid := FALSE;                             // 有效标志预置假 EN: preset the validity flag to false
nFaultCode := 0;                             // 故障码预置零 EN: preset the fault code to zero

// 段2｜非有限闸：五浮点入参全列
xFinAll := (rAccumLenM = rAccumLenM) AND ((rAccumLenM - rAccumLenM) = DL_WAC_Z)
        AND (rLineSpeedMpm = rLineSpeedMpm) AND ((rLineSpeedMpm - rLineSpeedMpm) = DL_WAC_Z)
        AND (rRollDiaMm = rRollDiaMm) AND ((rRollDiaMm - rRollDiaMm) = DL_WAC_Z)
        AND (rCoreDiaMm = rCoreDiaMm) AND ((rCoreDiaMm - rCoreDiaMm) = DL_WAC_Z)
        AND (rBufTimeMinS = rBufTimeMinS) AND ((rBufTimeMinS - rBufTimeMinS) = DL_WAC_Z);   // 五输入有限性 EN: the finiteness of all five inputs
IF NOT xFinAll THEN                                                                          // 非有限出口 EN: leave early on a non finite input
    nFaultCode := DL_WAC_C_BAD;                                                              // 非有限码 EN: the non finite code
    RETURN;                                                                                  // 早退 EN: return early
END_IF

// 段3｜域闸：储料长度与卷径非负、卷芯直径与线速度过分母下限
IF (rAccumLenM < DL_WAC_Z) OR (rRollDiaMm < DL_WAC_Z)
   OR (ABS(rCoreDiaMm) < DL_WAC_MIN) OR (ABS(rLineSpeedMpm) < DL_WAC_MIN) THEN
    nFaultCode := DL_WAC_C_RANGE;                                                            // 越域码 EN: the out of range code
    RETURN;                                                                                  // 早退 EN: return early
END_IF

// 段4｜主体：平均卷径 → 周长 → 圈数；线速度折每秒 → 缓冲时间（含饱和上限）
rMeanMm := (rRollDiaMm + rCoreDiaMm) / DL_WAC_TWO;                                           // 平均卷径 [mm] EN: the mean diameter
rMeanDiaM := rMeanMm / DL_WAC_K1000;                                                         // 平均卷径 [m] EN: the mean diameter in metres
rPerimM := DL_WAC_PI * rMeanDiaM;                                                            // 平均周长 [m] EN: the mean circumference
IF ABS(rPerimM) < DL_WAC_MIN THEN                                                            // 周长分母下限 EN: the circumference gate
    nFaultCode := DL_WAC_C_RANGE;                                                            // 越域码 EN: the out of range code
    RETURN;                                                                                  // 早退 EN: return early
END_IF
rWrap := rAccumLenM / rPerimM;                                                               // 折合圈数 [圈] EN: the equivalent wrap count
rSpeedMs := rLineSpeedMpm / DL_WAC_SECMIN;                                                   // 线速度 [m/s] EN: the line speed in metres per second
rTimeS := rAccumLenM / rSpeedMs;                                                             // 缓冲时间 [s] EN: the buffer time
IF rTimeS > DL_WAC_T_MAX THEN                                                                // 饱和上限（零速附近） EN: saturate near standstill
    rTimeS := DL_WAC_T_MAX;                                                                  // 饱和到上限 [s] EN: saturate to the upper bound
END_IF

// 段5｜结果复检与出口
IF (rWrap <> rWrap) OR (rTimeS <> rTimeS) OR (rWrap < DL_WAC_Z) OR (rTimeS < DL_WAC_Z) THEN   // 复检 EN: recheck the results
    nFaultCode := DL_WAC_C_RANGE;                                                            // 复检失败码 EN: the recheck failure code
    RETURN;                                                                                  // 早退，出口保持零哨兵 EN: return early with the zero sentinels
END_IF
rBufferTimeS := rTimeS;                                                                      // 缓冲时间出口 [s] EN: the buffer time output
rWrapCount := rWrap;                                                                         // 圈数出口 [圈] EN: the wrap count output
xBufferLow := rTimeS < rBufTimeMinS;                                                         // 缓冲不足判据（信息级） EN: the low buffer test, information class only
xValid := TRUE;                                                                              // 结果可信 EN: the results are valid
FC_DL_WebAccumulatorCapacityCalc := TRUE;                                                    // 返回真 EN: return true
END_FUNCTION

(* ---- FC_DL_WebGuideCamberCalc.st ---- *)
(*
  Component : FC_DL_WebGuideCamberCalc
  Category  : DL_Motion
  Function  : 镰刀弯曲率（三点弦高法）：camber = 8000 × h / L²，输出 mm/m 与等效曲率半径
  Complexity: C2
  开源溯源 : DLF 内部原创（R94 族模板派生）；参考语义来源见 SOURCE_HUNTING_MATRIX.md
  规则遵从 : R1-R16
  契约     : 输入 rChordMm 测量弦长（两基准点间距） [mm]、rSagittaMm 中点弦高（带符号） [mm]、
             rCamberMaxMmM 弯曲率工艺上限 [mm/m]；
             输出 rCamberMmM 带符号弯曲率 [mm/m]、rRadiusM 等效曲率半径 [m]、
             xCamberHigh 超上限（信息级）、xValid 有效标志、nFaultCode 故障码。
  边界     : 弦长须 >1.0E-6 [mm]；曲率半径 R = L²/(8h)，h 趋零时 R 趋于无穷，此时半径输出给 0 表示「直」；
             弯曲率 = 1000/R (R 以 mm 计时为 mm/m)，等价式 8000h/L²，符号随弦高；
             上限 1.0E4 [mm/m] 远小于 LREAL 上限，可表。
  码位     : 9801 输入非有限（故障级）；9802 弦长越域（故障级）。
*)
FUNCTION FC_DL_WebGuideCamberCalc : BOOL
VAR_INPUT
    rChordMm      : LREAL := 1000.0;  // 测量弦长 [mm] EN: the measured chord length
    rSagittaMm    : LREAL := 2.0;     // 中点弦高，正负表示弯曲方向 [mm] EN: the mid point sagitta, the sign carries the camber direction
    rCamberMaxMmM : LREAL := 5.0;     // 弯曲率工艺上限 [mm/m] EN: the technological upper bound of the camber rate
END_VAR
VAR_OUTPUT
    rCamberMmM  : LREAL;              // 带符号弯曲率 [mm/m] EN: the signed camber rate
    rRadiusM    : LREAL;              // 等效曲率半径，零表示直 [m] EN: the equivalent curvature radius, zero means straight
    xCamberHigh : BOOL;               // 超工艺上限（信息级） EN: above the technological limit, information class only
    xValid      : BOOL;               // 输出可信标志 EN: the outputs are valid
    nFaultCode  : INT;                // 0=无故障 9801=输入非有限 9802=弦长越域 EN: zero none, 9801 non finite, 9802 chord out of range
END_VAR
VAR
    xFinAll : BOOL;                   // 三输入同时有限 EN: all three inputs are finite
    rDen    : LREAL;                  // 分母 L²/8 [mm] EN: the divisor, the squared chord over eight
    rCam    : LREAL;                  // 弯曲率中间值 [mm/m] EN: the interim camber rate
    rRad    : LREAL;                  // 半径中间值 [m] EN: the interim radius
END_VAR
VAR CONSTANT
    DL_WGC_Z       : LREAL := 0.0;    // 浮点零常量 EN: the floating point zero constant
    DL_WGC_EIGHT   : LREAL := 8.0;    // 弦高法几何系数 EN: the geometric factor of the sagitta method
    DL_WGC_K1000   : LREAL := 1000.0; // 毫米转米系数 EN: the millimetre to metre factor
    DL_WGC_MIN     : LREAL := 1.0E-6; // 弦长与除数的下限 [mm] EN: the lower bound of the chord and the divisor
    DL_WGC_C_BAD   : INT := 9801;     // 输入非有限 EN: a non finite input
    DL_WGC_C_CHORD : INT := 9802;     // 弦长越域 EN: the chord is out of range
END_VAR

// 段1｜出口预置
FC_DL_WebGuideCamberCalc := FALSE;   // 返回值预置假 EN: preset the return value to false
rCamberMmM := DL_WGC_Z;               // 弯曲率预置零 [mm/m] EN: preset the camber rate to zero
rRadiusM := DL_WGC_Z;                 // 半径预置零 [m] EN: preset the radius to zero
xCamberHigh := FALSE;                 // 超限标志预置假 EN: preset the over camber flag to false
xValid := FALSE;                      // 有效标志预置假 EN: preset the validity flag to false
nFaultCode := 0;                      // 故障码预置零 EN: preset the fault code to zero

// 段2｜非有限闸：三输入全列（上限参与出口判据）
xFinAll := (rChordMm = rChordMm) AND ((rChordMm - rChordMm) = DL_WGC_Z)
        AND (rSagittaMm = rSagittaMm) AND ((rSagittaMm - rSagittaMm) = DL_WGC_Z)
        AND (rCamberMaxMmM = rCamberMaxMmM) AND ((rCamberMaxMmM - rCamberMaxMmM) = DL_WGC_Z);   // 三输入有限性 EN: the finiteness of all three inputs
IF NOT xFinAll THEN                                                                             // 非有限出口 EN: leave early on a non finite input
    nFaultCode := DL_WGC_C_BAD;                                                                 // 非有限码 EN: the non finite code
    RETURN;                                                                                     // 早退 EN: return early
END_IF

// 段3｜域闸：弦长必须足够大（分母 L²/8 直接依赖弦长）
rDen := (rChordMm * rChordMm) / DL_WGC_EIGHT;                                                   // 分母 L²/8 [mm] EN: the divisor
IF ABS(rDen) < DL_WGC_MIN THEN                                                                  // 分母下限 EN: the divisor magnitude gate
    nFaultCode := DL_WGC_C_CHORD;                                                               // 弦长越域码 EN: the chord code
    RETURN;                                                                                     // 早退 EN: return early
END_IF

// 段4｜主体：camber = h / (L²/8) × 1000 = 8000h/L²
rCam := (rSagittaMm / rDen) * DL_WGC_K1000;                                                     // 弯曲率 [mm/m]，符号随弦高 EN: the camber rate carrying the sagitta sign
IF rCam <> rCam THEN                                                                            // 结果复检 EN: recheck the result
    nFaultCode := DL_WGC_C_CHORD;                                                               // 复检失败码 EN: the recheck failure code
    RETURN;                                                                                     // 早退，出口保持零哨兵 EN: return early with the zero sentinels
END_IF

// 段5｜等效半径：弦高趋零时半径趋于无穷，统一给 0 表示直（不输出 Inf 污染上层）
IF ABS(rSagittaMm) < DL_WGC_MIN THEN                                                            // 近似直带 EN: the nearly straight band
    rRad := DL_WGC_Z;                                                                           // 半径给零表示直 [m] EN: give zero to mean straight
ELSE
    rRad := (rDen / rSagittaMm) / DL_WGC_K1000;                                                 // 半径 R = (L²/8)/h，由毫米折米 [m] EN: the radius folded to metres
END_IF

// 段6｜出口
rCamberMmM := rCam;                                                                             // 弯曲率出口 [mm/m] EN: the camber rate output
rRadiusM := rRad;                                                                               // 半径出口 [m] EN: the radius output
xCamberHigh := ABS(rCam) > rCamberMaxMmM;                                                       // 超限判据（信息级，双向均判） EN: the over camber test, information class, both directions
xValid := TRUE;                                                                                 // 结果可信 EN: the results are valid
FC_DL_WebGuideCamberCalc := TRUE;                                                               // 返回真 EN: return true
END_FUNCTION

(* ---- FC_DL_WebGuideDeadbandCalc.st ---- *)
(*
  Component : FC_DL_WebGuideDeadbandCalc
  Category  : DL_Motion
  Function  : 随线速度线性缩放的纠偏死区，含最小/最大钳位与速度上限保护
  Complexity: C2
  开源溯源 : DLF 内部原创（R94 族模板派生）；参考语义来源见 SOURCE_HUNTING_MATRIX.md
  规则遵从 : R1-R16
  契约     : 输入 rSpeedMpm 当前线速度 [m/min]、rSpeedRefMpm 速度归一化基准 [m/min]、
             rDeadbandMinMm 静止死区下限 [mm]、rDeadbandMaxMm 满速死区上限 [mm]；
             输出 rDeadbandMm 当前死区 [mm]、rSpeedRatio 速度比（未钳位） [-]、
             xSpeedCapped 速度比触上限、xValid 有效标志、nFaultCode 故障码。
  边界     : 速度比 = 当前速度 / 基准速度，基准速度须 >1.0E-6 [m/min]；速度比钳在 0~1（超基准速度不再放大死区，
             超速由运动层限速处理，本件不承担）；死区上下限须 0 ≤ min ≤ max。
  码位     : 9801 输入非有限（故障级）；9802 速度基准或死区上下限越域（故障级）。
*)
FUNCTION FC_DL_WebGuideDeadbandCalc : BOOL
VAR_INPUT
    rSpeedMpm      : LREAL := 100.0;  // 当前线速度 [m/min] EN: the current line speed
    rSpeedRefMpm   : LREAL := 200.0;  // 速度归一化基准 [m/min] EN: the reference speed used for normalisation
    rDeadbandMinMm : LREAL := 0.2;    // 静止死区下限 [mm] EN: the dead band at standstill
    rDeadbandMaxMm : LREAL := 1.0;    // 满速死区上限 [mm] EN: the dead band at the reference speed
END_VAR
VAR_OUTPUT
    rDeadbandMm  : LREAL;             // 当前纠偏死区 [mm] EN: the current guide dead band
    rSpeedRatio  : LREAL;             // 速度比（钳位后） [-] EN: the speed ratio after clamping
    xSpeedCapped : BOOL;              // 速度比触上限 EN: the speed ratio reached the upper bound
    xValid       : BOOL;              // 输出可信标志 EN: the outputs are valid
    nFaultCode   : INT;               // 0=无故障 9801=输入非有限 9802=基准或限值越域 EN: zero none, 9801 non finite, 9802 reference or limits out of range
END_VAR
VAR
    xFinAll : BOOL;                   // 四输入同时有限 EN: all four inputs are finite
    rRatio  : LREAL;                  // 速度比中间值 [-] EN: the interim speed ratio
    rRatioC : LREAL;                  // 钳位后速度比 [-] EN: the clamped speed ratio
    rDb     : LREAL;                  // 死区中间值 [mm] EN: the interim dead band
END_VAR
VAR CONSTANT
    DL_WGD_Z     : LREAL := 0.0;      // 浮点零常量 EN: the floating point zero constant
    DL_WGD_ONE   : LREAL := 1.0;      // 浮点壹常量 EN: the floating point one constant
    DL_WGD_MIN   : LREAL := 1.0E-6;   // 速度基准下限 [m/min] EN: the lower bound of the reference speed
    DL_WGD_C_BAD : INT := 9801;       // 输入非有限 EN: a non finite input
    DL_WGD_C_RANG: INT := 9802;       // 基准或限值越域 EN: the reference or the limits are out of range
END_VAR

// 段1｜出口预置
FC_DL_WebGuideDeadbandCalc := FALSE;   // 返回值预置假 EN: preset the return value to false
rDeadbandMm := DL_WGD_Z;               // 死区预置零 [mm] EN: preset the dead band to zero
rSpeedRatio := DL_WGD_Z;               // 速度比预置零 [-] EN: preset the speed ratio to zero
xSpeedCapped := FALSE;                 // 触限标志预置假 EN: preset the capped flag to false
xValid := FALSE;                       // 有效标志预置假 EN: preset the validity flag to false
nFaultCode := 0;                       // 故障码预置零 EN: preset the fault code to zero

// 段2｜非有限闸：四输入全列
xFinAll := (rSpeedMpm = rSpeedMpm) AND ((rSpeedMpm - rSpeedMpm) = DL_WGD_Z)
        AND (rSpeedRefMpm = rSpeedRefMpm) AND ((rSpeedRefMpm - rSpeedRefMpm) = DL_WGD_Z)
        AND (rDeadbandMinMm = rDeadbandMinMm) AND ((rDeadbandMinMm - rDeadbandMinMm) = DL_WGD_Z)
        AND (rDeadbandMaxMm = rDeadbandMaxMm) AND ((rDeadbandMaxMm - rDeadbandMaxMm) = DL_WGD_Z);   // 四输入有限性 EN: the finiteness of all four inputs
IF NOT xFinAll THEN                                                                                 // 非有限出口 EN: leave early on a non finite input
    nFaultCode := DL_WGD_C_BAD;                                                                     // 非有限码 EN: the non finite code
    RETURN;                                                                                         // 早退 EN: return early
END_IF

// 段3｜域闸：基准速度分母下限、速度非负、死区限值 0 ≤ min ≤ max
IF (ABS(rSpeedRefMpm) < DL_WGD_MIN) OR (rSpeedMpm < DL_WGD_Z)
   OR (rDeadbandMinMm < DL_WGD_Z) OR (rDeadbandMaxMm < rDeadbandMinMm) THEN
    nFaultCode := DL_WGD_C_RANG;                                                                    // 越域码 EN: the out of range code
    RETURN;                                                                                         // 早退 EN: return early
END_IF

// 段4｜主体：死区 = min + (max − min) × 速度比，速度比钳在 0~1
rRatio := rSpeedMpm / rSpeedRefMpm;                                                                 // 速度比 [-] EN: the speed ratio
rRatioC := rRatio;                                                                                  // 钳位工作副本 [-] EN: the working copy for clamping
IF rRatioC > DL_WGD_ONE THEN                                                                        // 上钳位 EN: clamp the upper bound
    rRatioC := DL_WGD_ONE;                                                                          // 钳到壹 [-] EN: clamp to one
    xSpeedCapped := TRUE;                                                                           // 置触限标志 EN: raise the capped flag
END_IF
IF rRatioC < DL_WGD_Z THEN                                                                          // 下钳位 EN: clamp the lower bound
    rRatioC := DL_WGD_Z;                                                                            // 钳到零 [-] EN: clamp to zero
END_IF
rDb := rDeadbandMinMm + (rDeadbandMaxMm - rDeadbandMinMm) * rRatioC;                                // 死区 [mm] EN: the dead band

// 段5｜出口：死区已在 [min,max] 内，另做一次非有限复检
IF (rDb <> rDb) OR (rDb < DL_WGD_Z) THEN                                                            // 复检 EN: recheck the result
    nFaultCode := DL_WGD_C_RANG;                                                                    // 复检失败码 EN: the recheck failure code
    RETURN;                                                                                         // 早退，出口保持零哨兵 EN: return early with the zero sentinels
END_IF
rDeadbandMm := rDb;                                                                                 // 死区出口 [mm] EN: the dead band output
rSpeedRatio := rRatioC;                                                                             // 速度比出口 [-] EN: the speed ratio output
xValid := TRUE;                                                                                     // 结果可信 EN: the results are valid
FC_DL_WebGuideDeadbandCalc := TRUE;                                                                 // 返回真 EN: return true
END_FUNCTION

(* ---- FC_DL_WebGuideRateLimitCalc.st ---- *)
(*
  Component : FC_DL_WebGuideRateLimitCalc
  Category  : DL_Motion
  Function  : 纠偏执行速率限幅：由剩余偏移量与最大加速度求允许速度 v = √(2·a·|e|)，并受最大速度钳制
  Complexity: C2
  开源溯源 : DLF 内部原创（R94 族模板派生）；参考语义来源见 SOURCE_HUNTING_MATRIX.md
  规则遵从 : R1-R16
  契约     : 输入 rOffsetMm 剩余偏移（带符号） [mm]、rAccelMmS2 允许最大加速度 [mm/s2]、
             rVmaxMmS 执行机构最大速度 [mm/s]、rDeadbandMm 纠偏死区 [mm]；
             输出 rVallowMmS 带符号允许速度 [mm/s]、rWithinDb 偏移在死区内、
             xLimited 触最大速度、xValid 有效标志、nFaultCode 故障码。
  边界     : 加速度与最大速度须 >0；偏移绝对值小于死区时允许速度给零（防抖）；
             速度符号随偏移符号，绝不取绝对值输出（符号即纠偏方向）；开方前乘子已证非负。
  码位     : 9801 输入非有限（故障级）；9802 加速度或最大速度越域（故障级）。
*)
FUNCTION FC_DL_WebGuideRateLimitCalc : BOOL
VAR_INPUT
    rOffsetMm   : LREAL := 1.0;      // 剩余带符号偏移 [mm] EN: the remaining signed offset
    rAccelMmS2  : LREAL := 50.0;     // 允许最大加速度 [mm/s2] EN: the allowed maximum acceleration
    rVmaxMmS    : LREAL := 20.0;     // 执行机构最大速度 [mm/s] EN: the maximum actuator velocity
    rDeadbandMm : LREAL := 0.2;      // 纠偏死区 [mm] EN: the guide dead band
END_VAR
VAR_OUTPUT
    rVallowMmS : LREAL;              // 带符号允许速度 [mm/s] EN: the signed allowed velocity
    rWithinDb  : BOOL;               // 偏移在死区内 EN: the offset is inside the dead band
    xLimited   : BOOL;               // 触最大速度 EN: the maximum velocity was reached
    xValid     : BOOL;               // 输出可信标志 EN: the outputs are valid
    nFaultCode : INT;                // 0=无故障 9801=输入非有限 9802=加速度或最大速度越域 EN: zero none, 9801 non finite, 9802 acceleration or maximum velocity out of range
END_VAR
VAR
    xFinAll : BOOL;                  // 四输入同时有限 EN: all four inputs are finite
    rAbsOff : LREAL;                 // 偏移绝对值 [mm] EN: the magnitude of the offset
    rEffOff : LREAL;                 // 扣死区后的有效偏移 [mm] EN: the effective offset after the dead band
    rVcalc  : LREAL;                 // 开方得到的限制速度 [mm/s] EN: the velocity limit from the square root
    rVout   : LREAL;                 // 允许速度幅值 [mm/s] EN: the allowed velocity magnitude
END_VAR
VAR CONSTANT
    DL_WRL_Z     : LREAL := 0.0;     // 浮点零常量 EN: the floating point zero constant
    DL_WRL_TWO   : LREAL := 2.0;     // 匀加速公式系数 EN: the uniform acceleration factor
    DL_WRL_C_BAD : INT := 9801;      // 输入非有限 EN: a non finite input
    DL_WRL_C_RANG: INT := 9802;      // 加速度或最大速度越域 EN: the acceleration or the maximum velocity is out of range
END_VAR

// 段1｜出口预置
FC_DL_WebGuideRateLimitCalc := FALSE;   // 返回值预置假 EN: preset the return value to false
rVallowMmS := DL_WRL_Z;                 // 允许速度预置零 [mm/s] EN: preset the allowed velocity to zero
rWithinDb := FALSE;                     // 死区标志预置假 EN: preset the dead band flag to false
xLimited := FALSE;                      // 触限标志预置假 EN: preset the limited flag to false
xValid := FALSE;                        // 有效标志预置假 EN: preset the validity flag to false
nFaultCode := 0;                        // 故障码预置零 EN: preset the fault code to zero

// 段2｜非有限闸：四输入全列（死区参与有效偏移，漏则防抖判据失效）
xFinAll := (rOffsetMm = rOffsetMm) AND ((rOffsetMm - rOffsetMm) = DL_WRL_Z)
        AND (rAccelMmS2 = rAccelMmS2) AND ((rAccelMmS2 - rAccelMmS2) = DL_WRL_Z)
        AND (rVmaxMmS = rVmaxMmS) AND ((rVmaxMmS - rVmaxMmS) = DL_WRL_Z)
        AND (rDeadbandMm = rDeadbandMm) AND ((rDeadbandMm - rDeadbandMm) = DL_WRL_Z);   // 四输入有限性 EN: the finiteness of all four inputs
IF NOT xFinAll THEN                                                                      // 非有限出口 EN: leave early on a non finite input
    nFaultCode := DL_WRL_C_BAD;                                                          // 非有限码 EN: the non finite code
    RETURN;                                                                              // 早退 EN: return early
END_IF

// 段3｜域闸：加速度与最大速度为正、死区非负
IF (rAccelMmS2 <= DL_WRL_Z) OR (rVmaxMmS <= DL_WRL_Z) OR (rDeadbandMm < DL_WRL_Z) THEN    // 域闸 EN: the domain gate
    nFaultCode := DL_WRL_C_RANG;                                                          // 越域码 EN: the out of range code
    RETURN;                                                                               // 早退 EN: return early
END_IF

// 段4｜主体：扣死区后按匀加速公式求限制速度，再与最大速度取小
rAbsOff := ABS(rOffsetMm);                                                                // 偏移绝对值 [mm] EN: the offset magnitude
rWithinDb := rAbsOff <= rDeadbandMm;                                                      // 死区判据 EN: the dead band test
rEffOff := rAbsOff - rDeadbandMm;                                                         // 有效偏移 [mm] EN: the effective offset
IF rWithinDb OR (rEffOff <= DL_WRL_Z) THEN                                                // 死区内或扣完无余量 EN: inside the band or nothing left
    rVout := DL_WRL_Z;                                                                    // 允许速度给零 [mm/s] EN: allow no motion
ELSE
    rVcalc := SQRT(DL_WRL_TWO * rAccelMmS2 * rEffOff);                                    // 匀加速限制速度，乘子已证正 [mm/s] EN: the square root limit, the operand is proven positive
    IF rVcalc > rVmaxMmS THEN                                                             // 与最大速度取小 EN: take the smaller bound
        rVout := rVmaxMmS;                                                                // 压到最大速度 [mm/s] EN: clamp to the maximum velocity
        xLimited := TRUE;                                                                 // 置触限标志 EN: raise the limited flag
    ELSE
        rVout := rVcalc;                                                                  // 采用公式值 [mm/s] EN: use the computed value
    END_IF
END_IF

// 段5｜出口：符号随偏移符号落定（R94 早退分支同样施加该变换）
IF rOffsetMm < DL_WRL_Z THEN                                                              // 偏移为负 EN: the offset is negative
    rVallowMmS := -rVout;                                                                 // 负向速度 [mm/s] EN: the negative velocity
ELSE
    rVallowMmS := rVout;                                                                  // 正向（含零）速度 [mm/s] EN: the positive velocity including zero
END_IF
xValid := TRUE;                                                                           // 结果可信 EN: the results are valid
FC_DL_WebGuideRateLimitCalc := TRUE;                                                      // 返回真 EN: return true
END_FUNCTION

(* ---- FC_DL_WebRewindTaperCalc.st ---- *)
(*
  Component : FC_DL_WebRewindTaperCalc
  Category  : DL_Motion
  Function  : 收卷锥度张力 T = T0 / (1 + taper × (D/D0 − 1))，卷径增大张力递减
  Complexity: C2
  开源溯源 : DLF 内部原创（R94 族模板派生）；参考语义来源见 SOURCE_HUNTING_MATRIX.md
  规则遵从 : R1-R16
  契约     : 输入 rT0N 初始（卷芯处）张力 [N]、rTaper 锥度系数 [-]、rDiaMm 当前卷径 [mm]、
             rCoreDiaMm 卷芯直径 D0 [mm]、rTaperMax 锥度系数上限 [-]；
             输出 rTensionN 当前张力 [N]、rDiaRatio 卷径比 D/D0 [-]、
             xTaperBad 锥度系数越域（信息级，按 0 处理并留痕）、xValid 有效标志、nFaultCode 故障码。
  边界     : 卷芯直径为分母须 >1.0E-6 [mm]；锥度分母 1 + taper×(ratio−1) 须 >1.0E-6（taper=−1 且卷径比
             恰为 2 时分母为零，属参数越域，判 9802）；初始张力须 ≥0；锥度系数按 [0, rTaperMax] 判域。
  码位     : 9801 输入非有限（故障级）；9802 卷芯直径或锥度分母越域（故障级）。
*)
FUNCTION FC_DL_WebRewindTaperCalc : BOOL
VAR_INPUT
    rT0N      : LREAL := 300.0;      // 卷芯处初始张力 [N] EN: the initial tension at the core
    rTaper    : LREAL := 0.3;        // 锥度系数 [-] EN: the taper coefficient
    rDiaMm    : LREAL := 600.0;      // 当前卷径 [mm] EN: the current roll diameter
    rCoreDiaMm: LREAL := 150.0;      // 卷芯直径 [mm] EN: the core diameter
    rTaperMax : LREAL := 1.0;        // 锥度系数上限 [-] EN: the upper bound of the taper coefficient
END_VAR
VAR_OUTPUT
    rTensionN : LREAL;               // 当前锥度张力 [N] EN: the current taper tension
    rDiaRatio : LREAL;               // 卷径比 D/D0 [-] EN: the diameter ratio
    xTaperBad : BOOL;                // 锥度系数越域（信息级） EN: the taper coefficient is out of range, information class only
    xValid    : BOOL;                // 输出可信标志 EN: the outputs are valid
    nFaultCode: INT;                 // 0=无故障 9801=输入非有限 9802=卷芯直径或锥度分母越域 EN: zero none, 9801 non finite, 9802 core diameter or taper divisor out of range
END_VAR
VAR
    xFinAll : BOOL;                  // 五输入同时有限 EN: all five inputs are finite
    rRatio  : LREAL;                 // 卷径比中间值 [-] EN: the interim diameter ratio
    rTaperU : LREAL;                 // 实际使用的锥度系数（越域时取零） [-] EN: the taper coefficient in use, zero when out of range
    rDen    : LREAL;                 // 锥度分母 [-] EN: the taper divisor
    rTens   : LREAL;                 // 张力中间值 [N] EN: the interim tension
END_VAR
VAR CONSTANT
    DL_WRT_Z     : LREAL := 0.0;     // 浮点零常量 EN: the floating point zero constant
    DL_WRT_ONE   : LREAL := 1.0;     // 浮点壹常量 EN: the floating point one constant
    DL_WRT_MIN   : LREAL := 1.0E-6;  // 分母绝对值下限 EN: the lower bound of the divisor magnitude
    DL_WRT_C_BAD : INT := 9801;      // 输入非有限 EN: a non finite input
    DL_WRT_C_DEN : INT := 9802;      // 卷芯直径或锥度分母越域 EN: the core diameter or the taper divisor is out of range
END_VAR

// 段1｜出口预置
FC_DL_WebRewindTaperCalc := FALSE;   // 返回值预置假 EN: preset the return value to false
rTensionN := DL_WRT_Z;               // 张力预置零 [N] EN: preset the tension to zero
rDiaRatio := DL_WRT_Z;               // 卷径比预置零 [-] EN: preset the diameter ratio to zero
xTaperBad := FALSE;                  // 锥度越域标志预置假 EN: preset the taper flag to false
xValid := FALSE;                     // 有效标志预置假 EN: preset the validity flag to false
nFaultCode := 0;                     // 故障码预置零 EN: preset the fault code to zero

// 段2｜非有限闸：五浮点入参全列
xFinAll := (rT0N = rT0N) AND ((rT0N - rT0N) = DL_WRT_Z)
        AND (rTaper = rTaper) AND ((rTaper - rTaper) = DL_WRT_Z)
        AND (rDiaMm = rDiaMm) AND ((rDiaMm - rDiaMm) = DL_WRT_Z)
        AND (rCoreDiaMm = rCoreDiaMm) AND ((rCoreDiaMm - rCoreDiaMm) = DL_WRT_Z)
        AND (rTaperMax = rTaperMax) AND ((rTaperMax - rTaperMax) = DL_WRT_Z);   // 五输入有限性 EN: the finiteness of all five inputs
IF NOT xFinAll THEN                                                            // 非有限出口 EN: leave early on a non finite input
    nFaultCode := DL_WRT_C_BAD;                                                // 非有限码 EN: the non finite code
    RETURN;                                                                    // 早退 EN: return early
END_IF

// 段3｜域闸：初始张力非负、卷芯直径为正、卷径非负、锥度上限非负
IF (rT0N < DL_WRT_Z) OR (rDiaMm < DL_WRT_Z) OR (rCoreDiaMm < DL_WRT_MIN) OR (rTaperMax < DL_WRT_Z) THEN
    nFaultCode := DL_WRT_C_DEN;                                                // 越域码 EN: the out of range code
    RETURN;                                                                    // 早退 EN: return early
END_IF

// 段4｜锥度系数域：越域按零（等效无锥度）处理并置信息级标志，不中断输出
IF (rTaper < DL_WRT_Z) OR (rTaper > rTaperMax) THEN                            // 锥度域判据 EN: the taper domain test
    rTaperU := DL_WRT_Z;                                                       // 越域取零（无锥度） [-] EN: fall back to zero
    xTaperBad := TRUE;                                                         // 置信息级标志 EN: raise the information class flag
ELSE
    rTaperU := rTaper;                                                         // 域内直接使用 [-] EN: use the coefficient as given
END_IF

// 段5｜主体：T = T0 / (1 + taper × (D/D0 − 1))
rRatio := rDiaMm / rCoreDiaMm;                                                 // 卷径比，分母已证正 [-] EN: the diameter ratio, the divisor is proven positive
rDen := DL_WRT_ONE + rTaperU * (rRatio - DL_WRT_ONE);                          // 锥度分母 [-] EN: the taper divisor
IF ABS(rDen) < DL_WRT_MIN THEN                                                 // 锥度分母下限 EN: the taper divisor gate
    nFaultCode := DL_WRT_C_DEN;                                                // 分母越域码 EN: the divisor code
    RETURN;                                                                    // 早退 EN: return early
END_IF
rTens := rT0N / rDen;                                                          // 锥度张力 [N] EN: the taper tension
IF (rTens <> rTens) OR (rTens < DL_WRT_Z) THEN                                 // 结果复检 EN: recheck the result
    nFaultCode := DL_WRT_C_DEN;                                                // 复检失败码 EN: the recheck failure code
    RETURN;                                                                    // 早退，出口保持零哨兵 EN: return early with the zero sentinels
END_IF

// 段6｜出口
rTensionN := rTens;                                                            // 张力出口 [N] EN: the tension output
rDiaRatio := rRatio;                                                           // 卷径比出口 [-] EN: the diameter ratio output
xValid := TRUE;                                                                // 结果可信 EN: the results are valid
FC_DL_WebRewindTaperCalc := TRUE;                                              // 返回真 EN: return true
END_FUNCTION

(* ---- FC_DL_WebSagCalc.st ---- *)
(*
  Component : FC_DL_WebSagCalc
  Category  : DL_Motion
  Function  : 卷材跨距垂度（悬链近似）sag = w·g·L²/(8T)，并给出垂度上限判定
  Complexity: C2
  开源溯源 : DLF 内部原创（R94 族模板派生）；参考语义来源见 SOURCE_HUNTING_MATRIX.md
  规则遵从 : R1-R16
  契约     : 输入 rSpanM 跨距（两支撑点间距） [m]、rLinearDensityKgM 卷材线密度 [kg/m]、
             rTensionN 带材张力 [N]、rSagMaxMm 垂度允许上限 [mm]；
             输出 rSagMm 垂度 [mm]、rSagRatioPct 垂度占跨距百分比 [%]、
             xSagHigh 超上限（信息级）、xValid 有效标志、nFaultCode 故障码。
  边界     : 张力为分母须 >1.0E-6 [N]（张力趋零垂度发散，悬链近似失效）；跨距与线密度须 ≥0；
             重力加速度取 9.80665 [m/s2]；垂度小于跨距的 1/8 时悬链近似误差 <2%，超出时仅作趋势参考。
  码位     : 9801 输入非有限（故障级）；9802 张力过小或跨距/线密度为负（故障级）。
*)
FUNCTION FC_DL_WebSagCalc : BOOL
VAR_INPUT
    rSpanM           : LREAL := 3.0;      // 跨距 [m] EN: the span between the two supports
    rLinearDensityKgM: LREAL := 0.5;      // 卷材线密度 [kg/m] EN: the linear density of the web
    rTensionN        : LREAL := 500.0;    // 带材张力 [N] EN: the web tension
    rSagMaxMm        : LREAL := 10.0;     // 垂度允许上限 [mm] EN: the allowed upper bound of the sag
END_VAR
VAR_OUTPUT
    rSagMm      : LREAL;                  // 垂度 [mm] EN: the sag in millimetres
    rSagRatioPct: LREAL;                  // 垂度占跨距百分比 [%] EN: the sag expressed as a percent of the span
    xSagHigh    : BOOL;                   // 超垂度上限（信息级） EN: above the sag limit, information class only
    xValid      : BOOL;                   // 输出可信标志 EN: the outputs are valid
    nFaultCode  : INT;                    // 0=无故障 9801=输入非有限 9802=张力过小或参数越域 EN: zero none, 9801 non finite, 9802 tension too small or parameters out of range
END_VAR
VAR
    xFinAll : BOOL;                       // 四输入同时有限 EN: all four inputs are finite
    rDen    : LREAL;                      // 分母 8T [N] EN: the divisor, eight times the tension
    rSagM   : LREAL;                      // 垂度中间值 [m] EN: the interim sag in metres
    rRatio  : LREAL;                      // 垂度比 [%] EN: the sag ratio in percent
END_VAR
VAR CONSTANT
    DL_WSC_Z       : LREAL := 0.0;        // 浮点零常量 EN: the floating point zero constant
    DL_WSC_G       : LREAL := 9.80665;    // 标准重力加速度 [m/s2] EN: the standard gravity acceleration
    DL_WSC_EIGHT   : LREAL := 8.0;        // 悬链近似几何系数 EN: the geometric factor of the catenary approximation
    DL_WSC_K1000   : LREAL := 1000.0;     // 米转毫米系数 EN: the metre to millimetre factor
    DL_WSC_HUNDRED : LREAL := 100.0;      // 百分数换算系数 EN: the percent conversion factor
    DL_WSC_MIN     : LREAL := 1.0E-6;     // 张力下限 [N] EN: the lower bound of the tension
    DL_WSC_C_BAD   : INT := 9801;         // 输入非有限 EN: a non finite input
    DL_WSC_C_RANGE : INT := 9802;         // 张力过小或参数越域 EN: the tension is too small or the parameters are out of range
END_VAR

// 段1｜出口预置
FC_DL_WebSagCalc := FALSE;   // 返回值预置假 EN: preset the return value to false
rSagMm := DL_WSC_Z;          // 垂度预置零 [mm] EN: preset the sag to zero
rSagRatioPct := DL_WSC_Z;    // 垂度比预置零 [%] EN: preset the sag ratio to zero
xSagHigh := FALSE;           // 超限标志预置假 EN: preset the over sag flag to false
xValid := FALSE;             // 有效标志预置假 EN: preset the validity flag to false
nFaultCode := 0;             // 故障码预置零 EN: preset the fault code to zero

// 段2｜非有限闸：四输入全列（上限参与出口判据）
xFinAll := (rSpanM = rSpanM) AND ((rSpanM - rSpanM) = DL_WSC_Z)
        AND (rLinearDensityKgM = rLinearDensityKgM) AND ((rLinearDensityKgM - rLinearDensityKgM) = DL_WSC_Z)
        AND (rTensionN = rTensionN) AND ((rTensionN - rTensionN) = DL_WSC_Z)
        AND (rSagMaxMm = rSagMaxMm) AND ((rSagMaxMm - rSagMaxMm) = DL_WSC_Z);   // 四输入有限性 EN: the finiteness of all four inputs
IF NOT xFinAll THEN                                                             // 非有限出口 EN: leave early on a non finite input
    nFaultCode := DL_WSC_C_BAD;                                                 // 非有限码 EN: the non finite code
    RETURN;                                                                     // 早退 EN: return early
END_IF

// 段3｜域闸：张力过分母下限、跨距与线密度非负
rDen := DL_WSC_EIGHT * rTensionN;                                              // 分母 8T [N] EN: the divisor
IF (ABS(rDen) < DL_WSC_MIN) OR (rSpanM < DL_WSC_Z) OR (rLinearDensityKgM < DL_WSC_Z) THEN
    nFaultCode := DL_WSC_C_RANGE;                                              // 越域码 EN: the out of range code
    RETURN;                                                                     // 早退 EN: return early
END_IF

// 段4｜主体：sag = w·g·L²/(8T)
rSagM := (rLinearDensityKgM * DL_WSC_G * rSpanM * rSpanM) / rDen;              // 垂度 [m] EN: the sag in metres
rSagMm := rSagM * DL_WSC_K1000;                                                // 垂度 [mm] EN: the sag in millimetres
IF (rSagMm <> rSagMm) OR (rSagMm < DL_WSC_Z) THEN                              // 结果复检 EN: recheck the result
    nFaultCode := DL_WSC_C_RANGE;                                              // 复检失败码 EN: the recheck failure code
    RETURN;                                                                     // 早退，出口保持零哨兵 EN: return early with the zero sentinels
END_IF

// 段5｜垂度占跨距百分比：跨距为零时不可比，给零
IF rSpanM > DL_WSC_MIN THEN                                                    // 跨距有效 EN: the span is usable
    rRatio := (rSagM / rSpanM) * DL_WSC_HUNDRED;                               // 垂度比 [%] EN: the sag ratio
ELSE
    rRatio := DL_WSC_Z;                                                        // 不可比给零 [%] EN: give zero when not comparable
END_IF

// 段6｜出口（垂度值在段4 已写入出口，此处只落定比值与超限判据，避免自赋值死语句）
rSagRatioPct := rRatio;                                                        // 垂度比出口 [%] EN: the sag ratio output
xSagHigh := rSagMm > rSagMaxMm;                                                // 超限判据（信息级） EN: the over sag test, information class only
xValid := TRUE;                                                               // 结果可信 EN: the results are valid
FC_DL_WebSagCalc := TRUE;                                                     // 返回真 EN: return true
END_FUNCTION

(* ---- FC_DL_WebSlitWidthCalc.st ---- *)
(*
  Component : FC_DL_WebSlitWidthCalc
  Category  : DL_Motion
  Function  : 分切宽度与边料核算：母卷宽 − n×成品宽，给出最大条数、边料总量与单边余量
  Complexity: C2
  开源溯源 : DLF 内部原创（R94 族模板派生）；参考语义来源见 SOURCE_HUNTING_MATRIX.md
  规则遵从 : R1-R16
  契约     : 输入 rMotherWidthMm 母卷有效宽度 [mm]、rProductWidthMm 成品宽度 [mm]、nSlits 计划分条数 [条]、
             rMinTrimPerSideMm 单边最小边料 [mm]；
             输出 nSlitsMax 理论最大条数 [条]、rTrimTotalMm 边料总量 [mm]、rTrimPerSideMm 单边边料 [mm]、
             xFeasible 方案可行（边料满足单边下限）、xValid 有效标志、nFaultCode 故障码。
  边界     : 成品宽度为分母须 >1.0E-6 [mm]；母卷宽与成品宽须 >0；分条数须 0~999；
             最大条数用向下取整（TRUNC），禁向上取整（多切一条即成品超宽，属不可返工缺陷）；
             边料均分时单边 = 总量/2，奇数宽度余量取小于 0.5 mm 的尾差并入单边下限判定。
  码位     : 9801 输入非有限（故障级）；9802 宽度越域或分条数越界（故障级）。
*)
FUNCTION FC_DL_WebSlitWidthCalc : BOOL
VAR_INPUT
    rMotherWidthMm   : LREAL := 1500.0;   // 母卷有效宽度 [mm] EN: the usable mother roll width
    rProductWidthMm  : LREAL := 300.0;    // 成品宽度 [mm] EN: the finished slit width
    nSlits           : INT := 4;          // 计划分条数 [条] EN: the planned number of slits
    rMinTrimPerSideMm: LREAL := 5.0;      // 单边最小边料 [mm] EN: the minimum trim per side
END_VAR
VAR_OUTPUT
    nSlitsMax     : INT;                  // 理论最大分条数 [条] EN: the theoretical maximum slit count
    rTrimTotalMm  : LREAL;                // 边料总量 [mm] EN: the total trim width
    rTrimPerSideMm: LREAL;                // 单边边料 [mm] EN: the trim per side
    xFeasible     : BOOL;                 // 方案可行 EN: the plan is feasible
    xValid        : BOOL;                 // 输出可信标志 EN: the outputs are valid
    nFaultCode    : INT;                  // 0=无故障 9801=输入非有限 9802=宽度或分条数越域 EN: zero none, 9801 non finite, 9802 width or slit count out of range
END_VAR
VAR
    xFinAll : BOOL;                       // 三个浮点入参有限 EN: the three floating inputs are finite
    rQuot   : LREAL;                      // 母卷宽与成品宽的商 [-] EN: the quotient of the mother width and the product width
    rTrim   : LREAL;                      // 边料总量中间值 [mm] EN: the interim total trim
    rSide   : LREAL;                      // 单边边料中间值 [mm] EN: the interim trim per side
    nMax    : INT;                        // 最大条数中间值 [条] EN: the interim maximum slit count
END_VAR
VAR CONSTANT
    DL_WSW_Z        : LREAL := 0.0;       // 浮点零常量 EN: the floating point zero constant
    DL_WSW_TWO      : LREAL := 2.0;       // 单边均分系数 EN: the per side splitting factor
    DL_WSW_SLIT_MAX : INT := 999;         // 分条数上限 [条] EN: the upper bound of the slit count
    DL_WSW_SLIT_MAXF: LREAL := 999.0;     // 分条数上限的实数值（转整前兜底） [条] EN: the real valued bound used before the integer conversion
    DL_WSW_MIN      : LREAL := 1.0E-6;    // 成品宽度下限 [mm] EN: the lower bound of the product width
    DL_WSW_C_BAD    : INT := 9801;        // 输入非有限 EN: a non finite input
    DL_WSW_C_RANGE  : INT := 9802;        // 宽度或分条数越域 EN: the width or the slit count is out of range
END_VAR

// 段1｜出口预置
FC_DL_WebSlitWidthCalc := FALSE;   // 返回值预置假 EN: preset the return value to false
nSlitsMax := 0;                    // 最大条数预置零 [条] EN: preset the maximum slit count to zero
rTrimTotalMm := DL_WSW_Z;          // 边料总量预置零 [mm] EN: preset the total trim to zero
rTrimPerSideMm := DL_WSW_Z;        // 单边边料预置零 [mm] EN: preset the trim per side to zero
xFeasible := FALSE;                // 可行标志预置假 EN: preset the feasibility flag to false
xValid := FALSE;                   // 有效标志预置假 EN: preset the validity flag to false
nFaultCode := 0;                   // 故障码预置零 EN: preset the fault code to zero

// 段2｜非有限闸：三浮点入参全列（单边下限参与可行性判据）
xFinAll := (rMotherWidthMm = rMotherWidthMm) AND ((rMotherWidthMm - rMotherWidthMm) = DL_WSW_Z)
        AND (rProductWidthMm = rProductWidthMm) AND ((rProductWidthMm - rProductWidthMm) = DL_WSW_Z)
        AND (rMinTrimPerSideMm = rMinTrimPerSideMm) AND ((rMinTrimPerSideMm - rMinTrimPerSideMm) = DL_WSW_Z);   // 三输入有限性 EN: the finiteness of all three inputs
IF NOT xFinAll THEN                                                                                           // 非有限出口 EN: leave early on a non finite input
    nFaultCode := DL_WSW_C_BAD;                                                                               // 非有限码 EN: the non finite code
    RETURN;                                                                                                   // 早退 EN: return early
END_IF

// 段3｜域闸：两宽度为正、成品宽过分母下限、单边下限非负、分条数 0~999
IF (rMotherWidthMm <= DL_WSW_Z) OR (ABS(rProductWidthMm) < DL_WSW_MIN)
   OR (rMinTrimPerSideMm < DL_WSW_Z) OR (nSlits < 0) OR (nSlits > DL_WSW_SLIT_MAX) THEN
    nFaultCode := DL_WSW_C_RANGE;                                                                             // 越域码 EN: the out of range code
    RETURN;                                                                                                   // 早退 EN: return early
END_IF

// 段4｜最大条数：向下取整（多切一条即成品超宽，故绝不上取整）
rQuot := rMotherWidthMm / rProductWidthMm;                                                                    // 商，分母已证正 [-] EN: the quotient, the divisor is proven positive
IF rQuot > DL_WSW_SLIT_MAXF THEN                                                                             // 实数上限兜底，防转 INT 溢出 EN: bound the real value before the integer conversion
    nMax := DL_WSW_SLIT_MAX;                                                                                 // 直接取上限 [条] EN: take the upper bound
ELSE
    nMax := LREAL_TO_INT(TRUNC(rQuot));                                                                      // 向下取整 [条] EN: truncate downwards
END_IF

// 段5｜按计划条数核算边料
rTrim := rMotherWidthMm - INT_TO_LREAL(nSlits) * rProductWidthMm;                                            // 边料总量 [mm] EN: the total trim
rSide := rTrim / DL_WSW_TWO;                                                                                 // 单边边料 [mm] EN: the trim per side
IF (rTrim <> rTrim) OR (rSide <> rSide) THEN                                                                  // 复检 EN: recheck
    nFaultCode := DL_WSW_C_RANGE;                                                                             // 复检失败码 EN: the recheck failure code
    RETURN;                                                                                                   // 早退，出口保持零哨兵 EN: return early with the zero sentinels
END_IF

// 段6｜出口：可行判据为「条数 ≥1 且 单边边料 ≥ 单边下限」
nSlitsMax := nMax;                                                                                           // 最大条数出口 [条] EN: the maximum slit count output
rTrimTotalMm := rTrim;                                                                                        // 边料总量出口 [mm] EN: the total trim output
rTrimPerSideMm := rSide;                                                                                      // 单边边料出口 [mm] EN: the trim per side output
xFeasible := (nSlits >= 1) AND (rSide >= rMinTrimPerSideMm);                                                  // 可行性判定 EN: the feasibility verdict
xValid := TRUE;                                                                                               // 结果可信 EN: the results are valid
FC_DL_WebSlitWidthCalc := TRUE;                                                                                // 返回真 EN: return true
END_FUNCTION

(* ---- FC_DL_WebTensionFromDancerCalc.st ---- *)
(*
  Component : FC_DL_WebTensionFromDancerCalc
  Category  : DL_Motion
  Function  : 浮辊位置折算张力 T = (F气缸 + k×Δx) / 走带股数，含零位与股数保护
  Complexity: C2
  开源溯源 : DLF 内部原创（R94 族模板派生）；参考语义来源见 SOURCE_HUNTING_MATRIX.md
  规则遵从 : R1-R16
  契约     : 输入 rDancerPosMm 浮辊实际位置 [mm]、rDancerZeroMm 浮辊零位（张力零点标定位置） [mm]、
             rStiffNPerMm 蓄能弹簧（或配重）等效刚度 [N/mm]、rCylForceN 气缸折算力 [N]、
             nStrandCount 走带股数 [股]；输出 rTensionN 单股张力 [N]、rDeflectMm 相对零位位移 [mm]、
             xNegTension 张力为负（信息级：带材松弛）、xValid 有效标志、nFaultCode 故障码。
  边界     : 股数须在 1~8 内（0 股为组态错误，判 9802）；弹簧刚度须 ≥0；位移可为负（浮辊下沉）；
             力平衡取「2 侧带材张力之和 = 气缸力 + 弹簧力」，故单股张力除以股数。
  码位     : 9801 输入非有限（故障级）；9802 股数或刚度越域（故障级）。
*)
FUNCTION FC_DL_WebTensionFromDancerCalc : BOOL
VAR_INPUT
    rDancerPosMm  : LREAL := 50.0;    // 浮辊实际位置 [mm] EN: the actual dancer position
    rDancerZeroMm : LREAL := 0.0;     // 浮辊张力零位标定值 [mm] EN: the calibrated dancer position at zero tension
    rStiffNPerMm  : LREAL := 0.5;     // 等效刚度（弹簧或配重折算） [N/mm] EN: the equivalent stiffness of the spring or the counterweight
    rCylForceN    : LREAL := 200.0;   // 气缸折算力（已扣自重） [N] EN: the cylinder force with the dead weight removed
    nStrandCount  : INT := 2;         // 走带股数 [股] EN: the number of web strands passing the dancer
END_VAR
VAR_OUTPUT
    rTensionN   : LREAL;              // 单股张力 [N] EN: the tension per strand
    rDeflectMm  : LREAL;              // 相对零位位移 [mm] EN: the displacement from the zero position
    xNegTension : BOOL;               // 张力为负（信息级，带材松弛） EN: a negative tension meaning a slack web, information class only
    xValid      : BOOL;               // 输出可信标志 EN: the outputs are valid
    nFaultCode  : INT;                // 0=无故障 9801=输入非有限 9802=股数或刚度越域 EN: zero none, 9801 non finite, 9802 strand count or stiffness out of range
END_VAR
VAR
    xFinAll : BOOL;                   // 四个浮点入参有限 EN: the four floating inputs are finite
    rDefl   : LREAL;                  // 位移中间值 [mm] EN: the interim displacement
    rForce  : LREAL;                  // 总力中间值 [N] EN: the interim total force
    rTens   : LREAL;                  // 单股张力中间值 [N] EN: the interim tension per strand
    rN      : LREAL;                  // 股数的实数形式 [股] EN: the strand count as a real number
END_VAR
VAR CONSTANT
    DL_WTD_Z      : LREAL := 0.0;     // 浮点零常量 EN: the floating point zero constant
    DL_WTD_STR_MAX: INT := 8;         // 股数上限 [股] EN: the upper bound of the strand count
    DL_WTD_C_BAD  : INT := 9801;      // 输入非有限 EN: a non finite input
    DL_WTD_C_RANGE: INT := 9802;      // 股数或刚度越域 EN: the strand count or the stiffness is out of range
END_VAR

// 段1｜出口预置
FC_DL_WebTensionFromDancerCalc := FALSE;   // 返回值预置假 EN: preset the return value to false
rTensionN := DL_WTD_Z;                      // 张力预置零 [N] EN: preset the tension to zero
rDeflectMm := DL_WTD_Z;                     // 位移预置零 [mm] EN: preset the displacement to zero
xNegTension := FALSE;                       // 负张力标志预置假 EN: preset the negative tension flag to false
xValid := FALSE;                            // 有效标志预置假 EN: preset the validity flag to false
nFaultCode := 0;                            // 故障码预置零 EN: preset the fault code to zero

// 段2｜非有限闸：四浮点入参全列
xFinAll := (rDancerPosMm = rDancerPosMm) AND ((rDancerPosMm - rDancerPosMm) = DL_WTD_Z)
        AND (rDancerZeroMm = rDancerZeroMm) AND ((rDancerZeroMm - rDancerZeroMm) = DL_WTD_Z)
        AND (rStiffNPerMm = rStiffNPerMm) AND ((rStiffNPerMm - rStiffNPerMm) = DL_WTD_Z)
        AND (rCylForceN = rCylForceN) AND ((rCylForceN - rCylForceN) = DL_WTD_Z);   // 四输入有限性 EN: the finiteness of all four inputs
IF NOT xFinAll THEN                                                                  // 非有限出口 EN: leave early on a non finite input
    nFaultCode := DL_WTD_C_BAD;                                                      // 非有限码 EN: the non finite code
    RETURN;                                                                          // 早退 EN: return early
END_IF

// 段3｜域闸：股数 1~8、刚度非负
IF (nStrandCount < 1) OR (nStrandCount > DL_WTD_STR_MAX) OR (rStiffNPerMm < DL_WTD_Z) THEN   // 股数与刚度闸 EN: the strand count and stiffness gate
    nFaultCode := DL_WTD_C_RANGE;                                                              // 越域码 EN: the out of range code
    RETURN;                                                                                    // 早退 EN: return early
END_IF

// 段4｜主体：总力 = 气缸力 + 刚度 × 位移；单股张力 = 总力 / 股数
rDefl := rDancerPosMm - rDancerZeroMm;                                                          // 相对零位位移 [mm] EN: the displacement from the zero position
rForce := rCylForceN + rStiffNPerMm * rDefl;                                                    // 总力 [N] EN: the total force
rN := INT_TO_LREAL(nStrandCount);                                                               // 股数实数化，已证 ≥1 [股] EN: the strand count as a real number, proven at least one
rTens := rForce / rN;                                                                           // 单股张力 [N] EN: the tension per strand

// 段5｜结果复检与出口
IF (rTens <> rTens) OR (rDefl <> rDefl) THEN                                                    // 复检：两路输出非有限 EN: recheck both outputs
    nFaultCode := DL_WTD_C_RANGE;                                                               // 复检失败码 EN: the recheck failure code
    RETURN;                                                                                     // 早退，出口保持零哨兵 EN: return early with the zero sentinels
END_IF
rDeflectMm := rDefl;                                                                            // 位移出口 [mm] EN: the displacement output
rTensionN := rTens;                                                                             // 张力出口 [N] EN: the tension output
xNegTension := rTens < DL_WTD_Z;                                                                // 负张力判据（信息级） EN: the negative tension test, information class only
xValid := TRUE;                                                                                 // 结果可信 EN: the results are valid
FC_DL_WebTensionFromDancerCalc := TRUE;                                                         // 返回真 EN: return true
END_FUNCTION

(* ---- FC_DL_WheelSlipRatioCalc.st ---- *)
// FC_DL_WheelSlipRatioCalc v1.0.0
// 开源溯源：clean-room 自研（族 DL_Motion，ST 生态实测 0 命中，无外部代码引入）
(*
  功能: 轮速滑移率 den = MAX(|v_veh|, 0.05)，s = (v_wheel − v_veh)/den，
        |s| > fSlipLimit 置打滑告警；den 下限保证静止时不除零。
  邻件/码位: 与 FC_DL_DiffDriveOdometryCalc 同属底盘状态件（打滑时里程计可信度下降）；
             fSlipLimit 非法取 0.2 缺省属信息级不置错；16#0002_9207 = 非有限拒收。
*)
FUNCTION FC_DL_WheelSlipRatioCalc : REAL
VAR_INPUT
    fWheelSpeed   : REAL := 0.0;    // 轮缘线速度 [m/s] / Wheel rim speed [m/s]
    fVehicleSpeed : REAL := 0.0;    // 车体车速 [m/s] / Vehicle body speed [m/s]
    fSlipLimit    : REAL := 0.2;    // 打滑阈值 [-]，<=0 取 0.2 / Slip threshold [-]
END_VAR
VAR_OUTPUT
    fSlipRatio : REAL;              // 滑移率 s [-]，驱动正 / Slip ratio [-]
    bSlipAlarm : BOOL;              // 打滑告警 [-] / Slip alarm flag
    bValid     : BOOL;              // 结果有效回执 [-] / Result validity receipt
    uErrorId   : UDINT;             // 事件码，0 = 无事件 / Event code
END_VAR
VAR
    fDen     : REAL := 0.0;         // 分母 MAX(|v_veh|, 0.05) [m/s] / Denominator [m/s]
    fLimitOk : REAL := 0.0;         // 生效阈值 [-] / Effective threshold [-]
    fAbsSlip : REAL := 0.0;         // 滑移率绝对值 [-] / Absolute slip ratio [-]
END_VAR
// 段 0：全路径出口安全缺省（滑移率零 + 告警清）/ Safe defaults
fSlipRatio := 0.0;              // 滑移率缺省零 / Slip ratio default zero
bSlipAlarm := FALSE;            // 告警预清 / Alarm preset clear
bValid := FALSE;                // 有效回执预清 / Validity preset clear
uErrorId := 16#0000;            // 事件码预清 / Event code preset clear
FC_DL_WheelSlipRatioCalc := 0.0;        // 返回值缺省零 / Return default zero
// 段 1：非有限闸（三入参全枚举）/ Non-finite gate over all inputs
IF (fWheelSpeed <> fWheelSpeed) OR (fVehicleSpeed <> fVehicleSpeed) OR (fSlipLimit <> fSlipLimit)
   OR (ABS(fWheelSpeed) >= 3.0E38) OR (ABS(fVehicleSpeed) >= 3.0E38) OR (ABS(fSlipLimit) >= 3.0E38) THEN
    uErrorId := 16#0002_9207;   // 入参非有限拒收 / Non-finite input reject
    RETURN;
END_IF
// 段 2：域闸（阈值非法取缺省 + 分母 0.05 硬下限）/ Domain gate, R4 divide-by-zero guard
fLimitOk := fSlipLimit;                                         // 阈值先直取 / Take as-is
IF fLimitOk <= 0.0 THEN
    fLimitOk := 0.2;                                            // 非法阈值取缺省 / Fallback to default
END_IF
fDen := ABS(fVehicleSpeed);                                     // 分母取车速绝对值 / Denominator initial
IF fDen < 0.05 THEN
    fDen := 0.05;                                               // 静止时保底防除零 / Static guard
END_IF
// 段 3：主计算（滑移率 + 告警判定）/ Main computation
fSlipRatio := (fWheelSpeed - fVehicleSpeed) / fDen;             // s = (vw − vv)/den / Slip ratio
fAbsSlip := ABS(fSlipRatio);                                    // 取绝对值 / Absolute value
IF fAbsSlip > fLimitOk THEN
    bSlipAlarm := TRUE;                                         // 超阈值告警 / Alarm above threshold
END_IF
// 段 4：出口闸（滑移率非有限复核）/ Outlet gate
IF (fSlipRatio <> fSlipRatio) OR (ABS(fSlipRatio) >= 3.0E38) THEN
    fSlipRatio := 0.0;          // 复核失败回缺省 / Fallback on recheck failure
    bSlipAlarm := FALSE;        // 复核失败清告警 / Clear alarm on recheck failure
    uErrorId := 16#0002_9207;   // 出口非有限拒收 / Output non-finite reject
    RETURN;
END_IF
bValid := TRUE;                 // 有效回执 / Validity receipt
FC_DL_WheelSlipRatioCalc := fSlipRatio; // 返回值镜像滑移率 / Return mirrors slip ratio
END_FUNCTION
